0.0, 0.0, 0.0, 0.0, 0.0, 0.0, 0.0, 0.0, 0.0, 0.0, 0.0, 0.0, 0.0, 0.0, 0.0, 0.0, 0.0, 0.0, 0.0, 0.0, 0.0, 0.0, 0.0, 0.0, 0.0, 0.0, 0.0, 0.0, 0.0, 0.0, 0.0, 0.0, 0.0, 0.0, 0.0, 0.0, 0.0, 0.0, 0.0, 0.0, 0.0, 0.0, 0.0, 0.0, 0.0, 0.0, 0.0, 0.0, 0.0, 0.0, 0.0, 0.0, 0.0, 0.0, 0.0, 0.0, 0.0, 0.0, 0.0, 0.0, 0.0, 0.0, 0.0, 0.0, 0.0, 0.0, -0.0, -0.0, -0.0, -0.0, -0.0, -0.0, -0.0, -0.0, -0.0, -0.0, -0.0, -0.0, -0.0, -0.0, -0.0, -0.0, -0.0, -0.0, -0.0, -0.0, -0.0, -0.0, -0.0, -0.0, -0.0, -0.0, -0.0, -0.0, -0.0, -0.0, -0.0, -0.0, -0.0, -0.0, -0.0, -0.0, -0.0, -0.0, -0.0, -0.0, -0.0, -0.0, -0.0, -0.0, -0.0, -0.0, -0.0, -0.0, -0.0, -0.0, -0.0, -0.0, -0.0, -0.0, -0.0, -0.0, -0.0, -0.0, -0.0, -0.0, -0.0, -0.0, -0.0, -0.0, -0.0, -0.0, -0.0, -0.0, -0.0, -0.0, -1.7756006070928429E-5, -1.955926027849794E-5, -2.1265642444599059E-5, -2.2878087249309936E-5, -2.4399475238503513E-5, -2.5832632877734329E-5, -2.7180332648224444E-5, -2.8445293182983732E-5, -2.9630179441154765E-5, -3.0737602918726609E-5, -3.1770121893815045E-5, -3.2730241704758869E-5, -3.3620415059333691E-5, -3.4443042373434618E-5, -3.5200472137629193E-5, -3.5895001310030509E-5, -3.652887573398812E-5, -3.7104290579141277E-5, -3.7623390804425058E-5, -3.808827164166491E-5, -3.8500979098439383E-5, -3.886351047893401E-5, -3.9177814921551905E-5, -3.9445793952087749E-5, -3.966930205131298E-5, -3.98501472358593E-5, -3.9990091651326829E-5, -4.0090852176581095E-5, -4.0154101038240283E-5, -4.0181466434390562E-5, -4.017453316660271E-5, -4.013484327935801E-5, -4.0063896706025282E-5, -3.9963151920563813E-5, -3.9834026594159355E-5, -3.9677898256031791E-5, -3.9496104957683613E-5, -3.9289945939888413E-5, -3.9060682301747689E-5, -3.8809537671172525E-5, -3.8537698876174604E-5, -3.8246316616377579E-5, -3.793650613418646E-5, -3.7609347885077623E-5, -3.7265888206497395E-5, -3.6907139984880808E-5, -3.6534083320325723E-5, -3.6147666188480321E-5, -3.5748805099224027E-5, -3.5338385751743129E-5, 0.0, 0.0, 0.0, 0.0, 0.0, 0.0, 0.0, 0.0, 0.0, 0.0, 0.0, 0.0, 0.0, 0.0, 0.0, 0.0, 0.0, 0.0, 0.0, 0.0, 0.0, 0.0, 0.0, 0.0, 0.0, 0.0, 0.0, 0.0, 0.0, 0.0, 0.0, 0.0, 0.0, 0.0, 0.0, 0.0, 0.0, 0.0, 0.0, 0.0, 0.0, 0.0, 0.0, 0.0, 0.0, 0.0, 0.0, 0.0, 0.0, 0.0, 0.0, 0.0, 0.0, 0.0, 0.0, 0.0, 0.0, 0.0, 0.0, 0.0, 0.0, 0.0, 0.0, 0.0, 0.0, 0.0, 0.0, 0.0, 0.0, 0.0, 1.7756006070928429E-5, 1.955926027849794E-5, 2.1265642444599059E-5, 2.2878087249309936E-5, 2.4399475238503513E-5, 2.5832632877734329E-5, 2.7180332648224444E-5, 2.8445293182983732E-5, 2.9630179441154765E-5, 3.0737602918726609E-5, 3.1770121893815045E-5, 3.2730241704758869E-5, 3.3620415059333691E-5, 3.4443042373434618E-5, 3.5200472137629193E-5, 3.5895001310030509E-5, 3.652887573398812E-5, 3.7104290579141277E-5, 3.7623390804425058E-5, 3.808827164166491E-5, 3.8500979098439383E-5, 3.886351047893401E-5, 3.9177814921551905E-5, 3.9445793952087749E-5, 3.966930205131298E-5, 3.98501472358593E-5, 3.9990091651326829E-5, 4.0090852176581095E-5, 4.0154101038240283E-5, 4.0181466434390562E-5, 4.017453316660271E-5, 4.013484327935801E-5, 4.0063896706025282E-5, 3.9963151920563813E-5, 3.9834026594159355E-5, 3.9677898256031791E-5, 3.9496104957683613E-5, 3.9289945939888413E-5, 3.9060682301747689E-5, 3.8809537671172525E-5, 3.8537698876174604E-5, 3.8246316616377579E-5, 3.793650613418646E-5, 3.7609347885077623E-5, 3.7265888206497395E-5, 3.6907139984880808E-5, 3.6534083320325723E-5, 3.6147666188480321E-5, 3.5748805099224027E-5, 3.5338385751743129E-5, 0.0, 0.0, 0.0, 0.0, -0.0, -0.0, -0.0, -0.0, -0.0, -0.0, -0.0, -0.0, -0.0, -0.0, -0.0, -0.0, -0.0, -0.0, -0.0, -0.0, -0.0, -0.0, -0.0, -0.0, -0.0, -0.0, -0.0, -0.0, -0.0, -0.0, -0.0, -0.0, -0.0, -0.0, -0.0, -0.0, -0.0, -0.0, -0.0, -0.0, -0.0, -0.0, -0.0, -0.0, -0.0, -0.0, -0.0, -0.0, -0.0, -0.0, -0.0, -0.0, -0.0, -0.0, -0.0, -0.0, -0.0, -0.0, -0.0, -0.0, -0.0, -0.0, -0.0, -0.0, -0.0, -0.0, -0.0, -0.0, -0.0, -0.0, -0.0, -0.0, -0.0, -0.0, -0.0, -0.0, -0.0, -0.0, -0.0, -0.0, -0.0, -0.0, -0.0, -0.0, -0.0, -0.0, -0.0, -0.0, -0.0, -0.0, -0.0, -0.0, -0.0, -0.0, -0.0, -0.0, -0.0, -0.0, -0.0, -0.0, -0.0, -0.0, -0.0, -0.0, -0.0, -0.0, -0.0, -0.0, -0.0, -0.0, -0.0, -0.0, -0.0, -0.0, -0.0, -0.0, -0.0, -0.0, -0.0, -0.0, -0.0, -0.0, -0.0, -0.0, 0.0, 0.0, 0.0, 0.0, 0.0, 0.0, 0.0, 0.0, 0.0, 0.0, 0.0, 0.0, 0.0, 0.0, 0.0, 0.0, 0.0, 0.0, 0.0, 0.0, 0.0, 0.0, 0.0, 0.0, 0.0, 0.0, 0.0, 0.0, 0.0, 0.0, 0.0, 0.0, 0.0, 0.0, 0.0, 0.0, 0.0, 0.0, 0.0, 0.0, 0.0, 0.0, 0.0, 0.0, 0.0, 0.0, 0.0, 0.0, 0.0, 0.0, 0.0, 0.0, 0.0, 0.0, 0.0, 0.0, 0.0, 0.0, 0.0, 0.0, 0.0, 0.0, 0.0, 0.0, 0.0, 0.0, 0.0, 0.0, 0.0, 0.0, 0.0, 0.0, 0.0, 0.0, 0.0, 0.0, 0.0, 0.0, 0.0, 0.0, 0.0, 0.0, 0.0, 0.0, 0.0, 0.0, 0.0, 0.0, 0.0, 0.0, 0.0, 0.0, 0.0, 0.0, 0.0, 0.0, 0.0, 0.0, 0.0, 0.0, 0.0, 0.0, 0.0, 0.0, 0.0, 0.0, 0.0, 0.0, 0.0, 0.0, 0.0, 0.0, 0.0, 0.0, 0.0, 0.0, 0.0, 0.0, 0.0, 0.0, 0.0, 0.0, 0.0, 0.0, -0.0, -0.0, -0.0, -0.0, -0.0, -0.0, -0.0, -0.0, -0.0, -0.0, -0.0, -0.0, -0.0, -0.0, -0.0, -0.0, -0.0, -0.0, -0.0, -0.0, -0.0, -0.0, -0.0, -0.0, -0.0, -0.0, -0.0, -0.0, -0.0, -0.0, -0.0, -0.0, -0.0, -0.0, -0.0, -0.0, -0.0, -0.0, -0.0, -0.0, -0.0, -0.0, -0.0, -0.0, -0.0, -0.0, -0.0, -0.0, -0.0, -0.0, -0.0, -0.0, -0.0, -0.0, -0.0, -0.0, -0.0, -0.0, -0.0, -0.0, -0.0, -0.0, -0.0, -0.0, -0.0, -0.0, -0.0, -0.0, -0.0, -0.0, -0.0, -1.7756006070928429E-5, -1.955926027849794E-5, -2.1265642444599059E-5, -2.2878087249309936E-5, -2.4399475238503513E-5, -2.5832632877734329E-5, -2.7180332648224444E-5, -2.8445293182983732E-5, -2.9630179441154765E-5, -3.0737602918726609E-5, -3.1770121893815045E-5, -3.2730241704758869E-5, -3.3620415059333691E-5, -3.4443042373434618E-5, -3.5200472137629193E-5, -3.5895001310030509E-5, -3.652887573398812E-5, -3.7104290579141277E-5, -3.7623390804425058E-5, -3.808827164166491E-5, -3.8500979098439383E-5, -3.886351047893401E-5, -3.9177814921551905E-5, -3.9445793952087749E-5, -3.966930205131298E-5, -3.98501472358593E-5, -3.9990091651326829E-5, -4.0090852176581095E-5, -4.0154101038240283E-5, -4.0181466434390562E-5, -4.017453316660271E-5, -4.013484327935801E-5, -4.0063896706025282E-5, -3.9963151920563813E-5, -3.9834026594159355E-5, -3.9677898256031791E-5, -3.9496104957683613E-5, -3.9289945939888413E-5, -3.9060682301747689E-5, -3.8809537671172525E-5, -3.8537698876174604E-5, -3.8246316616377579E-5, -3.793650613418646E-5, -3.7609347885077623E-5, -3.7265888206497395E-5, -3.6907139984880808E-5, -3.6534083320325723E-5, -3.6147666188480321E-5, -3.5748805099224027E-5, 0.0, 0.0, 0.0, 0.0, 0.0, 0.0, 0.0, 0.0, 0.0, 0.0, 0.0, 0.0, 0.0, 0.0, 0.0, 0.0, 0.0, 0.0, 0.0, 0.0, 0.0, 0.0, 0.0, 0.0, 0.0, 0.0, 0.0, 0.0, 0.0, 0.0, 0.0, 0.0, 0.0, 0.0, 0.0, 0.0, 0.0, 0.0, 0.0, 0.0, 0.0, 0.0, 0.0, 0.0, 0.0, 0.0, 0.0, 0.0, 0.0, 0.0, 0.0, 0.0, 0.0, 0.0, 0.0, 0.0, 0.0, 0.0, 0.0, 0.0, 0.0, 0.0, 0.0, 0.0, 0.0, 0.0, 0.0, 0.0, 0.0, 0.0, 0.0, 1.7756006070928429E-5, 1.955926027849794E-5, 2.1265642444599059E-5, 2.2878087249309936E-5, 2.4399475238503513E-5, 2.5832632877734329E-5, 2.7180332648224444E-5, 2.8445293182983732E-5, 2.9630179441154765E-5, 3.0737602918726609E-5, 3.1770121893815045E-5, 3.2730241704758869E-5, 3.3620415059333691E-5, 3.4443042373434618E-5, 3.5200472137629193E-5, 3.5895001310030509E-5, 3.652887573398812E-5, 3.7104290579141277E-5, 3.7623390804425058E-5, 3.808827164166491E-5, 3.8500979098439383E-5, 3.886351047893401E-5, 3.9177814921551905E-5, 3.9445793952087749E-5, 3.966930205131298E-5, 3.98501472358593E-5, 3.9990091651326829E-5, 4.0090852176581095E-5, 4.0154101038240283E-5, 4.0181466434390562E-5, 4.017453316660271E-5, 4.013484327935801E-5, 4.0063896706025282E-5, 3.9963151920563813E-5, 3.9834026594159355E-5, 3.9677898256031791E-5, 3.9496104957683613E-5, 3.9289945939888413E-5, 3.9060682301747689E-5, 3.8809537671172525E-5, 3.8537698876174604E-5, 3.8246316616377579E-5, 3.793650613418646E-5, 3.7609347885077623E-5, 3.7265888206497395E-5, 3.6907139984880808E-5, 3.6534083320325723E-5, 3.6147666188480321E-5, 3.5748805099224027E-5, 0.0, 0.0, 0.0, 0.0, -0.0, -0.0, -0.0, -0.0, -0.0, -0.0, -0.0, -0.0, -0.0, -0.0, -0.0, -0.0, -0.0, -0.0, -0.0, -0.0, -0.0, -0.0, -0.0, -0.0, -0.0, -0.0, -0.0, -0.0, -0.0, -0.0, -0.0, -0.0, -0.0, -0.0, -0.0, -0.0, -0.0, -0.0, -0.0, -0.0, -0.0, -0.0, -0.0, -0.0, -0.0, -0.0, -0.0, -0.0, -0.0, -0.0, -0.0, -0.0, -0.0, -0.0, -0.0, -0.0, -0.0, -0.0, -0.0, -0.0, -0.0, -0.0, -0.0, -0.0, -0.0, -0.0, -0.0, -0.0, -0.0, -0.0, -0.0, -0.0, -0.0, -0.0, -0.0, -0.0, -0.0, -0.0, -0.0, -0.0, -0.0, -0.0, -0.0, -0.0, -0.0, -0.0, -0.0, -0.0, -0.0, -0.0, -0.0, -0.0, -0.0, -0.0, -0.0, -0.0, -0.0, -0.0, -0.0, -0.0, -0.0, -0.0, -0.0, -0.0, -0.0, -0.0, -0.0, -0.0, -0.0, -0.0, -0.0, -0.0, -0.0, -0.0, -0.0, -0.0, -0.0, -0.0, -0.0, -0.0, -0.0, -0.0, -0.0, -0.0, 0.0, 0.0, 0.0, 0.0, 0.0, 0.0, 0.0, 0.0, 0.0, 0.0, 0.0, 0.0, 0.0, 0.0, 0.0, 0.0, 0.0, 0.0, 0.0, 0.0, 0.0, 0.0, 0.0, 0.0, 0.0, 0.0, 0.0, 0.0, 0.0, 0.0, 0.0, 0.0, 0.0, 0.0, 0.0, 0.0, 0.0, 0.0, 0.0, 0.0, 0.0, 0.0, 0.0, 0.0, 0.0, 0.0, 0.0, 0.0, 0.0, 0.0, 0.0, 0.0, 0.0, 0.0, 0.0, 0.0, 0.0, 0.0, 0.0, 0.0, 0.0, 0.0, 0.0, 0.0, 0.0, 0.0, 0.0, 0.0, 0.0, 0.0, 0.0, 0.0, 0.0, 0.0, 0.0, 0.0, 0.0, 0.0, 0.0, 0.0, 0.0, 0.0, 0.0, 0.0, 0.0, 0.0, 0.0, 0.0, 0.0, 0.0, 0.0, 0.0, 0.0, 0.0, 0.0, 0.0, 0.0, 0.0, 0.0, 0.0, 0.0, 0.0, 0.0, 0.0, 0.0, 0.0, 0.0, 0.0, 0.0, 0.0, 0.0, 0.0, 0.0, 0.0, 0.0, 0.0, 0.0, 0.0, 0.0, 0.0, 0.0, 0.0, 0.0, 0.0, -0.0, -0.0, -0.0, -0.0, -0.0, -0.0, -0.0, -0.0, -0.0, -0.0, -0.0, -0.0, -0.0, -0.0, -0.0, -0.0, -0.0, -0.0, -0.0, -0.0, -0.0, -0.0, -0.0, -0.0, -0.0, -0.0, -0.0, -0.0, -0.0, -0.0, -0.0, -0.0, -0.0, -0.0, -0.0, -0.0, -0.0, -0.0, -0.0, -0.0, -0.0, -0.0, -0.0, -0.0, -0.0, -0.0, -0.0, -0.0, -0.0, -0.0, -0.0, -0.0, -0.0, -0.0, -0.0, -0.0, -0.0, -0.0, -0.0, -0.0, -0.0, -0.0, -0.0, -0.0, -0.0, -0.0, -0.0, -0.0, -0.0, -0.0, -0.0, -0.0, -1.7756006070928429E-5, -1.955926027849794E-5, -2.1265642444599059E-5, -2.2878087249309936E-5, -2.4399475238503513E-5, -2.5832632877734329E-5, -2.7180332648224444E-5, -2.8445293182983732E-5, -2.9630179441154765E-5, -3.0737602918726609E-5, -3.1770121893815045E-5, -3.2730241704758869E-5, -3.3620415059333691E-5, -3.4443042373434618E-5, -3.5200472137629193E-5, -3.5895001310030509E-5, -3.652887573398812E-5, -3.7104290579141277E-5, -3.7623390804425058E-5, -3.808827164166491E-5, -3.8500979098439383E-5, -3.886351047893401E-5, -3.9177814921551905E-5, -3.9445793952087749E-5, -3.966930205131298E-5, -3.98501472358593E-5, -3.9990091651326829E-5, -4.0090852176581095E-5, -4.0154101038240283E-5, -4.0181466434390562E-5, -4.017453316660271E-5, -4.013484327935801E-5, -4.0063896706025282E-5, -3.9963151920563813E-5, -3.9834026594159355E-5, -3.9677898256031791E-5, -3.9496104957683613E-5, -3.9289945939888413E-5, -3.9060682301747689E-5, -3.8809537671172525E-5, -3.8537698876174604E-5, -3.8246316616377579E-5, -3.793650613418646E-5, -3.7609347885077623E-5, -3.7265888206497395E-5, -3.6907139984880808E-5, -3.6534083320325723E-5, -3.6147666188480321E-5, 0.0, 0.0, 0.0, 0.0, 0.0, 0.0, 0.0, 0.0, 0.0, 0.0, 0.0, 0.0, 0.0, 0.0, 0.0, 0.0, 0.0, 0.0, 0.0, 0.0, 0.0, 0.0, 0.0, 0.0, 0.0, 0.0, 0.0, 0.0, 0.0, 0.0, 0.0, 0.0, 0.0, 0.0, 0.0, 0.0, 0.0, 0.0, 0.0, 0.0, 0.0, 0.0, 0.0, 0.0, 0.0, 0.0, 0.0, 0.0, 0.0, 0.0, 0.0, 0.0, 0.0, 0.0, 0.0, 0.0, 0.0, 0.0, 0.0, 0.0, 0.0, 0.0, 0.0, 0.0, 0.0, 0.0, 0.0, 0.0, 0.0, 0.0, 0.0, 0.0, 1.7756006070928429E-5, 1.955926027849794E-5, 2.1265642444599059E-5, 2.2878087249309936E-5, 2.4399475238503513E-5, 2.5832632877734329E-5, 2.7180332648224444E-5, 2.8445293182983732E-5, 2.9630179441154765E-5, 3.0737602918726609E-5, 3.1770121893815045E-5, 3.2730241704758869E-5, 3.3620415059333691E-5, 3.4443042373434618E-5, 3.5200472137629193E-5, 3.5895001310030509E-5, 3.652887573398812E-5, 3.7104290579141277E-5, 3.7623390804425058E-5, 3.808827164166491E-5, 3.8500979098439383E-5, 3.886351047893401E-5, 3.9177814921551905E-5, 3.9445793952087749E-5, 3.966930205131298E-5, 3.98501472358593E-5, 3.9990091651326829E-5, 4.0090852176581095E-5, 4.0154101038240283E-5, 4.0181466434390562E-5, 4.017453316660271E-5, 4.013484327935801E-5, 4.0063896706025282E-5, 3.9963151920563813E-5, 3.9834026594159355E-5, 3.9677898256031791E-5, 3.9496104957683613E-5, 3.9289945939888413E-5, 3.9060682301747689E-5, 3.8809537671172525E-5, 3.8537698876174604E-5, 3.8246316616377579E-5, 3.793650613418646E-5, 3.7609347885077623E-5, 3.7265888206497395E-5, 3.6907139984880808E-5, 3.6534083320325723E-5, 3.6147666188480321E-5, 0.0, 0.0, 0.0, 0.0, -0.0, -0.0, -0.0, -0.0, -0.0, -0.0, -0.0, -0.0, -0.0, -0.0, -0.0, -0.0, -0.0, -0.0, -0.0, -0.0, -0.0, -0.0, -0.0, -0.0, -0.0, -0.0, -0.0, -0.0, -0.0, -0.0, -0.0, -0.0, -0.0, -0.0, -0.0, -0.0, -0.0, -0.0, -0.0, -0.0, -0.0, -0.0, -0.0, -0.0, -0.0, -0.0, -0.0, -0.0, -0.0, -0.0, -0.0, -0.0, -0.0, -0.0, -0.0, -0.0, -0.0, -0.0, -0.0, -0.0, -0.0, -0.0, -0.0, -0.0, -0.0, -0.0, -0.0, -0.0, -0.0, -0.0, -0.0, -0.0, -0.0, -0.0, -0.0, -0.0, -0.0, -0.0, -0.0, -0.0, -0.0, -0.0, -0.0, -0.0, -0.0, -0.0, -0.0, -0.0, -0.0, -0.0, -0.0, -0.0, -0.0, -0.0, -0.0, -0.0, -0.0, -0.0, -0.0, -0.0, -0.0, -0.0, -0.0, -0.0, -0.0, -0.0, -0.0, -0.0, -0.0, -0.0, -0.0, -0.0, -0.0, -0.0, -0.0, -0.0, -0.0, -0.0, -0.0, -0.0, -0.0, -0.0, -0.0, -0.0, 0.0, 0.0, 0.0, 0.0, 0.0, 0.0, 0.0, 0.0, 0.0, 0.0, 0.0, 0.0, 0.0, 0.0, 0.0, 0.0, 0.0, 0.0, 0.0, 0.0, 0.0, 0.0, 0.0, 0.0, 0.0, 0.0, 0.0, 0.0, 0.0, 0.0, 0.0, 0.0, 0.0, 0.0, 0.0, 0.0, 0.0, 0.0, 0.0, 0.0, 0.0, 0.0, 0.0, 0.0, 0.0, 0.0, 0.0, 0.0, 0.0, 0.0, 0.0, 0.0, 0.0, 0.0, 0.0, 0.0, 0.0, 0.0, 0.0, 0.0, 0.0, 0.0, 0.0, 0.0, 0.0, 0.0, 0.0, 0.0, 0.0, 0.0, 0.0, 0.0, 0.0, 0.0, 0.0, 0.0, 0.0, 0.0, 0.0, 0.0, 0.0, 0.0, 0.0, 0.0, 0.0, 0.0, 0.0, 0.0, 0.0, 0.0, 0.0, 0.0, 0.0, 0.0, 0.0, 0.0, 0.0, 0.0, 0.0, 0.0, 0.0, 0.0, 0.0, 0.0, 0.0, 0.0, 0.0, 0.0, 0.0, 0.0, 0.0, 0.0, 0.0, 0.0, 0.0, 0.0, 0.0, 0.0, 0.0, 0.0, 0.0, 0.0, 0.0, 0.0, -0.0, -0.0, -0.0, -0.0, -0.0, -0.0, -0.0, -0.0, -0.0, -0.0, -0.0, -0.0, -0.0, -0.0, -0.0, -0.0, -0.0, -0.0, -0.0, -0.0, -0.0, -0.0, -0.0, -0.0, -0.0, -0.0, -0.0, -0.0, -0.0, -0.0, -0.0, -0.0, -0.0, -0.0, -0.0, -0.0, -0.0, -0.0, -0.0, -0.0, -0.0, -0.0, -0.0, -0.0, -0.0, -0.0, -0.0, -0.0, -0.0, -0.0, -0.0, -0.0, -0.0, -0.0, -0.0, -0.0, -0.0, -0.0, -0.0, -0.0, -0.0, -0.0, -0.0, -0.0, -0.0, -0.0, -0.0, -0.0, -0.0, -0.0, -0.0, -0.0, -0.0, -1.7756006070928429E-5, -1.955926027849794E-5, -2.1265642444599059E-5, -2.2878087249309936E-5, -2.4399475238503513E-5, -2.5832632877734329E-5, -2.7180332648224444E-5, -2.8445293182983732E-5, -2.9630179441154765E-5, -3.0737602918726609E-5, -3.1770121893815045E-5, -3.2730241704758869E-5, -3.3620415059333691E-5, -3.4443042373434618E-5, -3.5200472137629193E-5, -3.5895001310030509E-5, -3.652887573398812E-5, -3.7104290579141277E-5, -3.7623390804425058E-5, -3.808827164166491E-5, -3.8500979098439383E-5, -3.886351047893401E-5, -3.9177814921551905E-5, -3.9445793952087749E-5, -3.966930205131298E-5, -3.98501472358593E-5, -3.9990091651326829E-5, -4.0090852176581095E-5, -4.0154101038240283E-5, -4.0181466434390562E-5, -4.017453316660271E-5, -4.013484327935801E-5, -4.0063896706025282E-5, -3.9963151920563813E-5, -3.9834026594159355E-5, -3.9677898256031791E-5, -3.9496104957683613E-5, -3.9289945939888413E-5, -3.9060682301747689E-5, -3.8809537671172525E-5, -3.8537698876174604E-5, -3.8246316616377579E-5, -3.793650613418646E-5, -3.7609347885077623E-5, -3.7265888206497395E-5, -3.6907139984880808E-5, -3.6534083320325723E-5, 0.0, 0.0, 0.0, 0.0, 0.0, 0.0, 0.0, 0.0, 0.0, 0.0, 0.0, 0.0, 0.0, 0.0, 0.0, 0.0, 0.0, 0.0, 0.0, 0.0, 0.0, 0.0, 0.0, 0.0, 0.0, 0.0, 0.0, 0.0, 0.0, 0.0, 0.0, 0.0, 0.0, 0.0, 0.0, 0.0, 0.0, 0.0, 0.0, 0.0, 0.0, 0.0, 0.0, 0.0, 0.0, 0.0, 0.0, 0.0, 0.0, 0.0, 0.0, 0.0, 0.0, 0.0, 0.0, 0.0, 0.0, 0.0, 0.0, 0.0, 0.0, 0.0, 0.0, 0.0, 0.0, 0.0, 0.0, 0.0, 0.0, 0.0, 0.0, 0.0, 0.0, 1.7756006070928429E-5, 1.955926027849794E-5, 2.1265642444599059E-5, 2.2878087249309936E-5, 2.4399475238503513E-5, 2.5832632877734329E-5, 2.7180332648224444E-5, 2.8445293182983732E-5, 2.9630179441154765E-5, 3.0737602918726609E-5, 3.1770121893815045E-5, 3.2730241704758869E-5, 3.3620415059333691E-5, 3.4443042373434618E-5, 3.5200472137629193E-5, 3.5895001310030509E-5, 3.652887573398812E-5, 3.7104290579141277E-5, 3.7623390804425058E-5, 3.808827164166491E-5, 3.8500979098439383E-5, 3.886351047893401E-5, 3.9177814921551905E-5, 3.9445793952087749E-5, 3.966930205131298E-5, 3.98501472358593E-5, 3.9990091651326829E-5, 4.0090852176581095E-5, 4.0154101038240283E-5, 4.0181466434390562E-5, 4.017453316660271E-5, 4.013484327935801E-5, 4.0063896706025282E-5, 3.9963151920563813E-5, 3.9834026594159355E-5, 3.9677898256031791E-5, 3.9496104957683613E-5, 3.9289945939888413E-5, 3.9060682301747689E-5, 3.8809537671172525E-5, 3.8537698876174604E-5, 3.8246316616377579E-5, 3.793650613418646E-5, 3.7609347885077623E-5, 3.7265888206497395E-5, 3.6907139984880808E-5, 3.6534083320325723E-5, 0.0, 0.0, 0.0, 0.0, -0.0, -0.0, -0.0, -0.0, -0.0, -0.0, -0.0, -0.0, -0.0, -0.0, -0.0, -0.0, -0.0, -0.0, -0.0, -0.0, -0.0, -0.0, -0.0, -0.0, -0.0, -0.0, -0.0, -0.0, -0.0, -0.0, -0.0, -0.0, -0.0, -0.0, -0.0, -0.0, -0.0, -0.0, -0.0, -0.0, -0.0, -0.0, -0.0, -0.0, -0.0, -0.0, -0.0, -0.0, -0.0, -0.0, -0.0, -0.0, -0.0, -0.0, -0.0, -0.0, -0.0, -0.0, -0.0, -0.0, -0.0, -0.0, -0.0, -0.0, -0.0, -0.0, -0.0, -0.0, -0.0, -0.0, -0.0, -0.0, -0.0, -0.0, -0.0, -0.0, -0.0, -0.0, -0.0, -0.0, -0.0, -0.0, -0.0, -0.0, -0.0, -0.0, -0.0, -0.0, -0.0, -0.0, -0.0, -0.0, -0.0, -0.0, -0.0, -0.0, -0.0, -0.0, -0.0, -0.0, -0.0, -0.0, -0.0, -0.0, -0.0, -0.0, -0.0, -0.0, -0.0, -0.0, -0.0, -0.0, -0.0, -0.0, -0.0, -0.0, -0.0, -0.0, -0.0, -0.0, -0.0, -0.0, -0.0, -0.0, 0.0, 0.0, 0.0, 0.0, 0.0, 0.0, 0.0, 0.0, 0.0, 0.0, 0.0, 0.0, 0.0, 0.0, 0.0, 0.0, 0.0, 0.0, 0.0, 0.0, 0.0, 0.0, 0.0, 0.0, 0.0, 0.0, 0.0, 0.0, 0.0, 0.0, 0.0, 0.0, 0.0, 0.0, 0.0, 0.0, 0.0, 0.0, 0.0, 0.0, 0.0, 0.0, 0.0, 0.0, 0.0, 0.0, 0.0, 0.0, 0.0, 0.0, 0.0, 0.0, 0.0, 0.0, 0.0, 0.0, 0.0, 0.0, 0.0, 0.0, 0.0, 0.0, 0.0, 0.0, 0.0, 0.0, 0.0, 0.0, 0.0, 0.0, 0.0, 0.0, 0.0, 0.0, 0.0, 0.0, 0.0, 0.0, 0.0, 0.0, 0.0, 0.0, 0.0, 0.0, 0.0, 0.0, 0.0, 0.0, 0.0, 0.0, 0.0, 0.0, 0.0, 0.0, 0.0, 0.0, 0.0, 0.0, 0.0, 0.0, 0.0, 0.0, 0.0, 0.0, 0.0, 0.0, 0.0, 0.0, 0.0, 0.0, 0.0, 0.0, 0.0, 0.0, 0.0, 0.0, 0.0, 0.0, 0.0, 0.0, 0.0, 0.0, 0.0, 0.0, -0.0, -0.0, -0.0, -0.0, -0.0, -0.0, -0.0, -0.0, -0.0, -0.0, -0.0, -0.0, -0.0, -0.0, -0.0, -0.0, -0.0, -0.0, -0.0, -0.0, -0.0, -0.0, -0.0, -0.0, -0.0, -0.0, -0.0, -0.0, -0.0, -0.0, -0.0, -0.0, -0.0, -0.0, -0.0, -0.0, -0.0, -0.0, -0.0, -0.0, -0.0, -0.0, -0.0, -0.0, -0.0, -0.0, -0.0, -0.0, -0.0, -0.0, -0.0, -0.0, -0.0, -0.0, -0.0, -0.0, -0.0, -0.0, -0.0, -0.0, -0.0, -0.0, -0.0, -0.0, -0.0, -0.0, -0.0, -0.0, -0.0, -0.0, -0.0, -0.0, -0.0, -0.0, -1.7756006070928429E-5, -1.955926027849794E-5, -2.1265642444599059E-5, -2.2878087249309936E-5, -2.4399475238503513E-5, -2.5832632877734329E-5, -2.7180332648224444E-5, -2.8445293182983732E-5, -2.9630179441154765E-5, -3.0737602918726609E-5, -3.1770121893815045E-5, -3.2730241704758869E-5, -3.3620415059333691E-5, -3.4443042373434618E-5, -3.5200472137629193E-5, -3.5895001310030509E-5, -3.652887573398812E-5, -3.7104290579141277E-5, -3.7623390804425058E-5, -3.808827164166491E-5, -3.8500979098439383E-5, -3.886351047893401E-5, -3.9177814921551905E-5, -3.9445793952087749E-5, -3.966930205131298E-5, -3.98501472358593E-5, -3.9990091651326829E-5, -4.0090852176581095E-5, -4.0154101038240283E-5, -4.0181466434390562E-5, -4.017453316660271E-5, -4.013484327935801E-5, -4.0063896706025282E-5, -3.9963151920563813E-5, -3.9834026594159355E-5, -3.9677898256031791E-5, -3.9496104957683613E-5, -3.9289945939888413E-5, -3.9060682301747689E-5, -3.8809537671172525E-5, -3.8537698876174604E-5, -3.8246316616377579E-5, -3.793650613418646E-5, -3.7609347885077623E-5, -3.7265888206497395E-5, -3.6907139984880808E-5, 0.0, 0.0, 0.0, 0.0, 0.0, 0.0, 0.0, 0.0, 0.0, 0.0, 0.0, 0.0, 0.0, 0.0, 0.0, 0.0, 0.0, 0.0, 0.0, 0.0, 0.0, 0.0, 0.0, 0.0, 0.0, 0.0, 0.0, 0.0, 0.0, 0.0, 0.0, 0.0, 0.0, 0.0, 0.0, 0.0, 0.0, 0.0, 0.0, 0.0, 0.0, 0.0, 0.0, 0.0, 0.0, 0.0, 0.0, 0.0, 0.0, 0.0, 0.0, 0.0, 0.0, 0.0, 0.0, 0.0, 0.0, 0.0, 0.0, 0.0, 0.0, 0.0, 0.0, 0.0, 0.0, 0.0, 0.0, 0.0, 0.0, 0.0, 0.0, 0.0, 0.0, 0.0, 1.7756006070928429E-5, 1.955926027849794E-5, 2.1265642444599059E-5, 2.2878087249309936E-5, 2.4399475238503513E-5, 2.5832632877734329E-5, 2.7180332648224444E-5, 2.8445293182983732E-5, 2.9630179441154765E-5, 3.0737602918726609E-5, 3.1770121893815045E-5, 3.2730241704758869E-5, 3.3620415059333691E-5, 3.4443042373434618E-5, 3.5200472137629193E-5, 3.5895001310030509E-5, 3.652887573398812E-5, 3.7104290579141277E-5, 3.7623390804425058E-5, 3.808827164166491E-5, 3.8500979098439383E-5, 3.886351047893401E-5, 3.9177814921551905E-5, 3.9445793952087749E-5, 3.966930205131298E-5, 3.98501472358593E-5, 3.9990091651326829E-5, 4.0090852176581095E-5, 4.0154101038240283E-5, 4.0181466434390562E-5, 4.017453316660271E-5, 4.013484327935801E-5, 4.0063896706025282E-5, 3.9963151920563813E-5, 3.9834026594159355E-5, 3.9677898256031791E-5, 3.9496104957683613E-5, 3.9289945939888413E-5, 3.9060682301747689E-5, 3.8809537671172525E-5, 3.8537698876174604E-5, 3.8246316616377579E-5, 3.793650613418646E-5, 3.7609347885077623E-5, 3.7265888206497395E-5, 3.6907139984880808E-5, 0.0, 0.0, 0.0, 0.0, -0.0, -0.0, -0.0, -0.0, -0.0, -0.0, -0.0, -0.0, -0.0, -0.0, -0.0, -0.0, -0.0, -0.0, -0.0, -0.0, -0.0, -0.0, -0.0, -0.0, -0.0, -0.0, -0.0, -0.0, -0.0, -0.0, -0.0, -0.0, -0.0, -0.0, -0.0, -0.0, -0.0, -0.0, -0.0, -0.0, -0.0, -0.0, -0.0, -0.0, -0.0, -0.0, -0.0, -0.0, -0.0, -0.0, -0.0, -0.0, -0.0, -0.0, -0.0, -0.0, -0.0, -0.0, -0.0, -0.0, -0.0, -0.0, -0.0, -0.0, -0.0, -0.0, -0.0, -0.0, -0.0, -0.0, -0.0, -0.0, -0.0, -0.0, -0.0, -0.0, -0.0, -0.0, -0.0, -0.0, -0.0, -0.0, -0.0, -0.0, -0.0, -0.0, -0.0, -0.0, -0.0, -0.0, -0.0, -0.0, -0.0, -0.0, -0.0, -0.0, -0.0, -0.0, -0.0, -0.0, -0.0, -0.0, -0.0, -0.0, -0.0, -0.0, -0.0, -0.0, -0.0, -0.0, -0.0, -0.0, -0.0, -0.0, -0.0, -0.0, -0.0, -0.0, -0.0, -0.0, -0.0, -0.0, -0.0, -0.0, 0.0, 0.0, 0.0, 0.0, 0.0, 0.0, 0.0, 0.0, 0.0, 0.0, 0.0, 0.0, 0.0, 0.0, 0.0, 0.0, 0.0, 0.0, 0.0, 0.0, 0.0, 0.0, 0.0, 0.0, 0.0, 0.0, 0.0, 0.0, 0.0, 0.0, 0.0, 0.0, 0.0, 0.0, 0.0, 0.0, 0.0, 0.0, 0.0, 0.0, 0.0, 0.0, 0.0, 0.0, 0.0, 0.0, 0.0, 0.0, 0.0, 0.0, 0.0, 0.0, 0.0, 0.0, 0.0, 0.0, 0.0, 0.0, 0.0, 0.0, 0.0, 0.0, 0.0, 0.0, 0.0, 0.0, 0.0, 0.0, 0.0, 0.0, 0.0, 0.0, 0.0, 0.0, 0.0, 0.0, 0.0, 0.0, 0.0, 0.0, 0.0, 0.0, 0.0, 0.0, 0.0, 0.0, 0.0, 0.0, 0.0, 0.0, 0.0, 0.0, 0.0, 0.0, 0.0, 0.0, 0.0, 0.0, 0.0, 0.0, 0.0, 0.0, 0.0, 0.0, 0.0, 0.0, 0.0, 0.0, 0.0, 0.0, 0.0, 0.0, 0.0, 0.0, 0.0, 0.0, 0.0, 0.0, 0.0, 0.0, 0.0, 0.0, 0.0, 0.0, -0.0, -0.0, -0.0, -0.0, -0.0, -0.0, -0.0, -0.0, -0.0, -0.0, -0.0, -0.0, -0.0, -0.0, -0.0, -0.0, -0.0, -0.0, -0.0, -0.0, -0.0, -0.0, -0.0, -0.0, -0.0, -0.0, -0.0, -0.0, -0.0, -0.0, -0.0, -0.0, -0.0, -0.0, -0.0, -0.0, -0.0, -0.0, -0.0, -0.0, -0.0, -0.0, -0.0, -0.0, -0.0, -0.0, -0.0, -0.0, -0.0, -0.0, -0.0, -0.0, -0.0, -0.0, -0.0, -0.0, -0.0, -0.0, -0.0, -0.0, -0.0, -0.0, -0.0, -0.0, -0.0, -0.0, -0.0, -0.0, -0.0, -0.0, -0.0, -0.0, -0.0, -0.0, -0.0, -1.7756006070928429E-5, -1.955926027849794E-5, -2.1265642444599059E-5, -2.2878087249309936E-5, -2.4399475238503513E-5, -2.5832632877734329E-5, -2.7180332648224444E-5, -2.8445293182983732E-5, -2.9630179441154765E-5, -3.0737602918726609E-5, -3.1770121893815045E-5, -3.2730241704758869E-5, -3.3620415059333691E-5, -3.4443042373434618E-5, -3.5200472137629193E-5, -3.5895001310030509E-5, -3.652887573398812E-5, -3.7104290579141277E-5, -3.7623390804425058E-5, -3.808827164166491E-5, -3.8500979098439383E-5, -3.886351047893401E-5, -3.9177814921551905E-5, -3.9445793952087749E-5, -3.966930205131298E-5, -3.98501472358593E-5, -3.9990091651326829E-5, -4.0090852176581095E-5, -4.0154101038240283E-5, -4.0181466434390562E-5, -4.017453316660271E-5, -4.013484327935801E-5, -4.0063896706025282E-5, -3.9963151920563813E-5, -3.9834026594159355E-5, -3.9677898256031791E-5, -3.9496104957683613E-5, -3.9289945939888413E-5, -3.9060682301747689E-5, -3.8809537671172525E-5, -3.8537698876174604E-5, -3.8246316616377579E-5, -3.793650613418646E-5, -3.7609347885077623E-5, -3.7265888206497395E-5, 0.0, 0.0, 0.0, 0.0, 0.0, 0.0, 0.0, 0.0, 0.0, 0.0, 0.0, 0.0, 0.0, 0.0, 0.0, 0.0, 0.0, 0.0, 0.0, 0.0, 0.0, 0.0, 0.0, 0.0, 0.0, 0.0, 0.0, 0.0, 0.0, 0.0, 0.0, 0.0, 0.0, 0.0, 0.0, 0.0, 0.0, 0.0, 0.0, 0.0, 0.0, 0.0, 0.0, 0.0, 0.0, 0.0, 0.0, 0.0, 0.0, 0.0, 0.0, 0.0, 0.0, 0.0, 0.0, 0.0, 0.0, 0.0, 0.0, 0.0, 0.0, 0.0, 0.0, 0.0, 0.0, 0.0, 0.0, 0.0, 0.0, 0.0, 0.0, 0.0, 0.0, 0.0, 0.0, 1.7756006070928429E-5, 1.955926027849794E-5, 2.1265642444599059E-5, 2.2878087249309936E-5, 2.4399475238503513E-5, 2.5832632877734329E-5, 2.7180332648224444E-5, 2.8445293182983732E-5, 2.9630179441154765E-5, 3.0737602918726609E-5, 3.1770121893815045E-5, 3.2730241704758869E-5, 3.3620415059333691E-5, 3.4443042373434618E-5, 3.5200472137629193E-5, 3.5895001310030509E-5, 3.652887573398812E-5, 3.7104290579141277E-5, 3.7623390804425058E-5, 3.808827164166491E-5, 3.8500979098439383E-5, 3.886351047893401E-5, 3.9177814921551905E-5, 3.9445793952087749E-5, 3.966930205131298E-5, 3.98501472358593E-5, 3.9990091651326829E-5, 4.0090852176581095E-5, 4.0154101038240283E-5, 4.0181466434390562E-5, 4.017453316660271E-5, 4.013484327935801E-5, 4.0063896706025282E-5, 3.9963151920563813E-5, 3.9834026594159355E-5, 3.9677898256031791E-5, 3.9496104957683613E-5, 3.9289945939888413E-5, 3.9060682301747689E-5, 3.8809537671172525E-5, 3.8537698876174604E-5, 3.8246316616377579E-5, 3.793650613418646E-5, 3.7609347885077623E-5, 3.7265888206497395E-5, 0.0, 0.0, 0.0, 0.0, -0.0, -0.0, -0.0, -0.0, -0.0, -0.0, -0.0, -0.0, -0.0, -0.0, -0.0, -0.0, -0.0, -0.0, -0.0, -0.0, -0.0, -0.0, -0.0, -0.0, -0.0, -0.0, -0.0, -0.0, -0.0, -0.0, -0.0, -0.0, -0.0, -0.0, -0.0, -0.0, -0.0, -0.0, -0.0, -0.0, -0.0, -0.0, -0.0, -0.0, -0.0, -0.0, -0.0, -0.0, -0.0, -0.0, -0.0, -0.0, -0.0, -0.0, -0.0, -0.0, -0.0, -0.0, -0.0, -0.0, -0.0, -0.0, -0.0, -0.0, -0.0, -0.0, -0.0, -0.0, -0.0, -0.0, -0.0, -0.0, -0.0, -0.0, -0.0, -0.0, -0.0, -0.0, -0.0, -0.0, -0.0, -0.0, -0.0, -0.0, -0.0, -0.0, -0.0, -0.0, -0.0, -0.0, -0.0, -0.0, -0.0, -0.0, -0.0, -0.0, -0.0, -0.0, -0.0, -0.0, -0.0, -0.0, -0.0, -0.0, -0.0, -0.0, -0.0, -0.0, -0.0, -0.0, -0.0, -0.0, -0.0, -0.0, -0.0, -0.0, -0.0, -0.0, -0.0, -0.0, -0.0, -0.0, -0.0, -0.0, 0.0, 0.0, 0.0, 0.0, 0.0, 0.0, 0.0, 0.0, 0.0, 0.0, 0.0, 0.0, 0.0, 0.0, 0.0, 0.0, 0.0, 0.0, 0.0, 0.0, 0.0, 0.0, 0.0, 0.0, 0.0, 0.0, 0.0, 0.0, 0.0, 0.0, 0.0, 0.0, 0.0, 0.0, 0.0, 0.0, 0.0, 0.0, 0.0, 0.0, 0.0, 0.0, 0.0, 0.0, 0.0, 0.0, 0.0, 0.0, 0.0, 0.0, 0.0, 0.0, 0.0, 0.0, 0.0, 0.0, 0.0, 0.0, 0.0, 0.0, 0.0, 0.0, 0.0, 0.0, 0.0, 0.0, 0.0, 0.0, 0.0, 0.0, 0.0, 0.0, 0.0, 0.0, 0.0, 0.0, 0.0, 0.0, 0.0, 0.0, 0.0, 0.0, 0.0, 0.0, 0.0, 0.0, 0.0, 0.0, 0.0, 0.0, 0.0, 0.0, 0.0, 0.0, 0.0, 0.0, 0.0, 0.0, 0.0, 0.0, 0.0, 0.0, 0.0, 0.0, 0.0, 0.0, 0.0, 0.0, 0.0, 0.0, 0.0, 0.0, 0.0, 0.0, 0.0, 0.0, 0.0, 0.0, 0.0, 0.0, 0.0, 0.0, 0.0, 0.0, -0.0, -0.0, -0.0, -0.0, -0.0, -0.0, -0.0, -0.0, -0.0, -0.0, -0.0, -0.0, -0.0, -0.0, -0.0, -0.0, -0.0, -0.0, -0.0, -0.0, -0.0, -0.0, -0.0, -0.0, -0.0, -0.0, -0.0, -0.0, -0.0, -0.0, -0.0, -0.0, -0.0, -0.0, -0.0, -0.0, -0.0, -0.0, -0.0, -0.0, -0.0, -0.0, -0.0, -0.0, -0.0, -0.0, -0.0, -0.0, -0.0, -0.0, -0.0, -0.0, -0.0, -0.0, -0.0, -0.0, -0.0, -0.0, -0.0, -0.0, -0.0, -0.0, -0.0, -0.0, -0.0, -0.0, -0.0, -0.0, -0.0, -0.0, -0.0, -0.0, -0.0, -0.0, -0.0, -0.0, -1.7756006070928429E-5, -1.955926027849794E-5, -2.1265642444599059E-5, -2.2878087249309936E-5, -2.4399475238503513E-5, -2.5832632877734329E-5, -2.7180332648224444E-5, -2.8445293182983732E-5, -2.9630179441154765E-5, -3.0737602918726609E-5, -3.1770121893815045E-5, -3.2730241704758869E-5, -3.3620415059333691E-5, -3.4443042373434618E-5, -3.5200472137629193E-5, -3.5895001310030509E-5, -3.652887573398812E-5, -3.7104290579141277E-5, -3.7623390804425058E-5, -3.808827164166491E-5, -3.8500979098439383E-5, -3.886351047893401E-5, -3.9177814921551905E-5, -3.9445793952087749E-5, -3.966930205131298E-5, -3.98501472358593E-5, -3.9990091651326829E-5, -4.0090852176581095E-5, -4.0154101038240283E-5, -4.0181466434390562E-5, -4.017453316660271E-5, -4.013484327935801E-5, -4.0063896706025282E-5, -3.9963151920563813E-5, -3.9834026594159355E-5, -3.9677898256031791E-5, -3.9496104957683613E-5, -3.9289945939888413E-5, -3.9060682301747689E-5, -3.8809537671172525E-5, -3.8537698876174604E-5, -3.8246316616377579E-5, -3.793650613418646E-5, -3.7609347885077623E-5, 0.0, 0.0, 0.0, 0.0, 0.0, 0.0, 0.0, 0.0, 0.0, 0.0, 0.0, 0.0, 0.0, 0.0, 0.0, 0.0, 0.0, 0.0, 0.0, 0.0, 0.0, 0.0, 0.0, 0.0, 0.0, 0.0, 0.0, 0.0, 0.0, 0.0, 0.0, 0.0, 0.0, 0.0, 0.0, 0.0, 0.0, 0.0, 0.0, 0.0, 0.0, 0.0, 0.0, 0.0, 0.0, 0.0, 0.0, 0.0, 0.0, 0.0, 0.0, 0.0, 0.0, 0.0, 0.0, 0.0, 0.0, 0.0, 0.0, 0.0, 0.0, 0.0, 0.0, 0.0, 0.0, 0.0, 0.0, 0.0, 0.0, 0.0, 0.0, 0.0, 0.0, 0.0, 0.0, 0.0, 1.7756006070928429E-5, 1.955926027849794E-5, 2.1265642444599059E-5, 2.2878087249309936E-5, 2.4399475238503513E-5, 2.5832632877734329E-5, 2.7180332648224444E-5, 2.8445293182983732E-5, 2.9630179441154765E-5, 3.0737602918726609E-5, 3.1770121893815045E-5, 3.2730241704758869E-5, 3.3620415059333691E-5, 3.4443042373434618E-5, 3.5200472137629193E-5, 3.5895001310030509E-5, 3.652887573398812E-5, 3.7104290579141277E-5, 3.7623390804425058E-5, 3.808827164166491E-5, 3.8500979098439383E-5, 3.886351047893401E-5, 3.9177814921551905E-5, 3.9445793952087749E-5, 3.966930205131298E-5, 3.98501472358593E-5, 3.9990091651326829E-5, 4.0090852176581095E-5, 4.0154101038240283E-5, 4.0181466434390562E-5, 4.017453316660271E-5, 4.013484327935801E-5, 4.0063896706025282E-5, 3.9963151920563813E-5, 3.9834026594159355E-5, 3.9677898256031791E-5, 3.9496104957683613E-5, 3.9289945939888413E-5, 3.9060682301747689E-5, 3.8809537671172525E-5, 3.8537698876174604E-5, 3.8246316616377579E-5, 3.793650613418646E-5, 3.7609347885077623E-5, 0.0, 0.0, 0.0, 0.0, -0.0, -0.0, -0.0, -0.0, -0.0, -0.0, -0.0, -0.0, -0.0, -0.0, -0.0, -0.0, -0.0, -0.0, -0.0, -0.0, -0.0, -0.0, -0.0, -0.0, -0.0, -0.0, -0.0, -0.0, -0.0, -0.0, -0.0, -0.0, -0.0, -0.0, -0.0, -0.0, -0.0, -0.0, -0.0, -0.0, -0.0, -0.0, -0.0, -0.0, -0.0, -0.0, -0.0, -0.0, -0.0, -0.0, -0.0, -0.0, -0.0, -0.0, -0.0, -0.0, -0.0, -0.0, -0.0, -0.0, -0.0, -0.0, -0.0, -0.0, -0.0, -0.0, -0.0, -0.0, -0.0, -0.0, -0.0, -0.0, -0.0, -0.0, -0.0, -0.0, -0.0, -0.0, -0.0, -0.0, -0.0, -0.0, -0.0, -0.0, -0.0, -0.0, -0.0, -0.0, -0.0, -0.0, -0.0, -0.0, -0.0, -0.0, -0.0, -0.0, -0.0, -0.0, -0.0, -0.0, -0.0, -0.0, -0.0, -0.0, -0.0, -0.0, -0.0, -0.0, -0.0, -0.0, -0.0, -0.0, -0.0, -0.0, -0.0, -0.0, -0.0, -0.0, -0.0, -0.0, -0.0, -0.0, -0.0, -0.0, 0.0, 0.0, 0.0, 0.0, 0.0, 0.0, 0.0, 0.0, 0.0, 0.0, 0.0, 0.0, 0.0, 0.0, 0.0, 0.0, 0.0, 0.0, 0.0, 0.0, 0.0, 0.0, 0.0, 0.0, 0.0, 0.0, 0.0, 0.0, 0.0, 0.0, 0.0, 0.0, 0.0, 0.0, 0.0, 0.0, 0.0, 0.0, 0.0, 0.0, 0.0, 0.0, 0.0, 0.0, 0.0, 0.0, 0.0, 0.0, 0.0, 0.0, 0.0, 0.0, 0.0, 0.0, 0.0, 0.0, 0.0, 0.0, 0.0, 0.0, 0.0, 0.0, 0.0, 0.0, 0.0, 0.0, 0.0, 0.0, 0.0, 0.0, 0.0, 0.0, 0.0, 0.0, 0.0, 0.0, 0.0, 0.0, 0.0, 0.0, 0.0, 0.0, 0.0, 0.0, 0.0, 0.0, 0.0, 0.0, 0.0, 0.0, 0.0, 0.0, 0.0, 0.0, 0.0, 0.0, 0.0, 0.0, 0.0, 0.0, 0.0, 0.0, 0.0, 0.0, 0.0, 0.0, 0.0, 0.0, 0.0, 0.0, 0.0, 0.0, 0.0, 0.0, 0.0, 0.0, 0.0, 0.0, 0.0, 0.0, 0.0, 0.0, 0.0, 0.0, -0.0, -0.0, -0.0, -0.0, -0.0, -0.0, -0.0, -0.0, -0.0, -0.0, -0.0, -0.0, -0.0, -0.0, -0.0, -0.0, -0.0, -0.0, -0.0, -0.0, -0.0, -0.0, -0.0, -0.0, -0.0, -0.0, -0.0, -0.0, -0.0, -0.0, -0.0, -0.0, -0.0, -0.0, -0.0, -0.0, -0.0, -0.0, -0.0, -0.0, -0.0, -0.0, -0.0, -0.0, -0.0, -0.0, -0.0, -0.0, -0.0, -0.0, -0.0, -0.0, -0.0, -0.0, -0.0, -0.0, -0.0, -0.0, -0.0, -0.0, -0.0, -0.0, -0.0, -0.0, -0.0, -0.0, -0.0, -0.0, -0.0, -0.0, -0.0, -0.0, -0.0, -0.0, -0.0, -0.0, -0.0, -1.7756006070928429E-5, -1.955926027849794E-5, -2.1265642444599059E-5, -2.2878087249309936E-5, -2.4399475238503513E-5, -2.5832632877734329E-5, -2.7180332648224444E-5, -2.8445293182983732E-5, -2.9630179441154765E-5, -3.0737602918726609E-5, -3.1770121893815045E-5, -3.2730241704758869E-5, -3.3620415059333691E-5, -3.4443042373434618E-5, -3.5200472137629193E-5, -3.5895001310030509E-5, -3.652887573398812E-5, -3.7104290579141277E-5, -3.7623390804425058E-5, -3.808827164166491E-5, -3.8500979098439383E-5, -3.886351047893401E-5, -3.9177814921551905E-5, -3.9445793952087749E-5, -3.966930205131298E-5, -3.98501472358593E-5, -3.9990091651326829E-5, -4.0090852176581095E-5, -4.0154101038240283E-5, -4.0181466434390562E-5, -4.017453316660271E-5, -4.013484327935801E-5, -4.0063896706025282E-5, -3.9963151920563813E-5, -3.9834026594159355E-5, -3.9677898256031791E-5, -3.9496104957683613E-5, -3.9289945939888413E-5, -3.9060682301747689E-5, -3.8809537671172525E-5, -3.8537698876174604E-5, -3.8246316616377579E-5, -3.793650613418646E-5, 0.0, 0.0, 0.0, 0.0, 0.0, 0.0, 0.0, 0.0, 0.0, 0.0, 0.0, 0.0, 0.0, 0.0, 0.0, 0.0, 0.0, 0.0, 0.0, 0.0, 0.0, 0.0, 0.0, 0.0, 0.0, 0.0, 0.0, 0.0, 0.0, 0.0, 0.0, 0.0, 0.0, 0.0, 0.0, 0.0, 0.0, 0.0, 0.0, 0.0, 0.0, 0.0, 0.0, 0.0, 0.0, 0.0, 0.0, 0.0, 0.0, 0.0, 0.0, 0.0, 0.0, 0.0, 0.0, 0.0, 0.0, 0.0, 0.0, 0.0, 0.0, 0.0, 0.0, 0.0, 0.0, 0.0, 0.0, 0.0, 0.0, 0.0, 0.0, 0.0, 0.0, 0.0, 0.0, 0.0, 0.0, 1.7756006070928429E-5, 1.955926027849794E-5, 2.1265642444599059E-5, 2.2878087249309936E-5, 2.4399475238503513E-5, 2.5832632877734329E-5, 2.7180332648224444E-5, 2.8445293182983732E-5, 2.9630179441154765E-5, 3.0737602918726609E-5, 3.1770121893815045E-5, 3.2730241704758869E-5, 3.3620415059333691E-5, 3.4443042373434618E-5, 3.5200472137629193E-5, 3.5895001310030509E-5, 3.652887573398812E-5, 3.7104290579141277E-5, 3.7623390804425058E-5, 3.808827164166491E-5, 3.8500979098439383E-5, 3.886351047893401E-5, 3.9177814921551905E-5, 3.9445793952087749E-5, 3.966930205131298E-5, 3.98501472358593E-5, 3.9990091651326829E-5, 4.0090852176581095E-5, 4.0154101038240283E-5, 4.0181466434390562E-5, 4.017453316660271E-5, 4.013484327935801E-5, 4.0063896706025282E-5, 3.9963151920563813E-5, 3.9834026594159355E-5, 3.9677898256031791E-5, 3.9496104957683613E-5, 3.9289945939888413E-5, 3.9060682301747689E-5, 3.8809537671172525E-5, 3.8537698876174604E-5, 3.8246316616377579E-5, 3.793650613418646E-5, 0.0, 0.0, 0.0, 0.0, -0.0, -0.0, -0.0, -0.0, -0.0, -0.0, -0.0, -0.0, -0.0, -0.0, -0.0, -0.0, -0.0, -0.0, -0.0, -0.0, -0.0, -0.0, -0.0, -0.0, -0.0, -0.0, -0.0, -0.0, -0.0, -0.0, -0.0, -0.0, -0.0, -0.0, -0.0, -0.0, -0.0, -0.0, -0.0, -0.0, -0.0, -0.0, -0.0, -0.0, -0.0, -0.0, -0.0, -0.0, -0.0, -0.0, -0.0, -0.0, -0.0, -0.0, -0.0, -0.0, -0.0, -0.0, -0.0, -0.0, -0.0, -0.0, -0.0, -0.0, -0.0, -0.0, -0.0, -0.0, -0.0, -0.0, -0.0, -0.0, -0.0, -0.0, -0.0, -0.0, -0.0, -0.0, -0.0, -0.0, -0.0, -0.0, -0.0, -0.0, -0.0, -0.0, -0.0, -0.0, -0.0, -0.0, -0.0, -0.0, -0.0, -0.0, -0.0, -0.0, -0.0, -0.0, -0.0, -0.0, -0.0, -0.0, -0.0, -0.0, -0.0, -0.0, -0.0, -0.0, -0.0, -0.0, -0.0, -0.0, -0.0, -0.0, -0.0, -0.0, -0.0, -0.0, -0.0, -0.0, -0.0, -0.0, -0.0, -0.0, 0.0, 0.0, 0.0, 0.0, 0.0, 0.0, 0.0, 0.0, 0.0, 0.0, 0.0, 0.0, 0.0, 0.0, 0.0, 0.0, 0.0, 0.0, 0.0, 0.0, 0.0, 0.0, 0.0, 0.0, 0.0, 0.0, 0.0, 0.0, 0.0, 0.0, 0.0, 0.0, 0.0, 0.0, 0.0, 0.0, 0.0, 0.0, 0.0, 0.0, 0.0, 0.0, 0.0, 0.0, 0.0, 0.0, 0.0, 0.0, 0.0, 0.0, 0.0, 0.0, 0.0, 0.0, 0.0, 0.0, 0.0, 0.0, 0.0, 0.0, 0.0, 0.0, 0.0, 0.0, 0.0, 0.0, 0.0, 0.0, 0.0, 0.0, 0.0, 0.0, 0.0, 0.0, 0.0, 0.0, 0.0, 0.0, 0.0, 0.0, 0.0, 0.0, 0.0, 0.0, 0.0, 0.0, 0.0, 0.0, 0.0, 0.0, 0.0, 0.0, 0.0, 0.0, 0.0, 0.0, 0.0, 0.0, 0.0, 0.0, 0.0, 0.0, 0.0, 0.0, 0.0, 0.0, 0.0, 0.0, 0.0, 0.0, 0.0, 0.0, 0.0, 0.0, 0.0, 0.0, 0.0, 0.0, 0.0, 0.0, 0.0, 0.0, 0.0, 0.0, -0.0, -0.0, -0.0, -0.0, -0.0, -0.0, -0.0, -0.0, -0.0, -0.0, -0.0, -0.0, -0.0, -0.0, -0.0, -0.0, -0.0, -0.0, -0.0, -0.0, -0.0, -0.0, -0.0, -0.0, -0.0, -0.0, -0.0, -0.0, -0.0, -0.0, -0.0, -0.0, -0.0, -0.0, -0.0, -0.0, -0.0, -0.0, -0.0, -0.0, -0.0, -0.0, -0.0, -0.0, -0.0, -0.0, -0.0, -0.0, -0.0, -0.0, -0.0, -0.0, -0.0, -0.0, -0.0, -0.0, -0.0, -0.0, -0.0, -0.0, -0.0, -0.0, -0.0, -0.0, -0.0, -0.0, -0.0, -0.0, -0.0, -0.0, -0.0, -0.0, -0.0, -0.0, -0.0, -0.0, -0.0, -0.0, -1.7756006070928429E-5, -1.955926027849794E-5, -2.1265642444599059E-5, -2.2878087249309936E-5, -2.4399475238503513E-5, -2.5832632877734329E-5, -2.7180332648224444E-5, -2.8445293182983732E-5, -2.9630179441154765E-5, -3.0737602918726609E-5, -3.1770121893815045E-5, -3.2730241704758869E-5, -3.3620415059333691E-5, -3.4443042373434618E-5, -3.5200472137629193E-5, -3.5895001310030509E-5, -3.652887573398812E-5, -3.7104290579141277E-5, -3.7623390804425058E-5, -3.808827164166491E-5, -3.8500979098439383E-5, -3.886351047893401E-5, -3.9177814921551905E-5, -3.9445793952087749E-5, -3.966930205131298E-5, -3.98501472358593E-5, -3.9990091651326829E-5, -4.0090852176581095E-5, -4.0154101038240283E-5, -4.0181466434390562E-5, -4.017453316660271E-5, -4.013484327935801E-5, -4.0063896706025282E-5, -3.9963151920563813E-5, -3.9834026594159355E-5, -3.9677898256031791E-5, -3.9496104957683613E-5, -3.9289945939888413E-5, -3.9060682301747689E-5, -3.8809537671172525E-5, -3.8537698876174604E-5, -3.8246316616377579E-5, 0.0, 0.0, 0.0, 0.0, 0.0, 0.0, 0.0, 0.0, 0.0, 0.0, 0.0, 0.0, 0.0, 0.0, 0.0, 0.0, 0.0, 0.0, 0.0, 0.0, 0.0, 0.0, 0.0, 0.0, 0.0, 0.0, 0.0, 0.0, 0.0, 0.0, 0.0, 0.0, 0.0, 0.0, 0.0, 0.0, 0.0, 0.0, 0.0, 0.0, 0.0, 0.0, 0.0, 0.0, 0.0, 0.0, 0.0, 0.0, 0.0, 0.0, 0.0, 0.0, 0.0, 0.0, 0.0, 0.0, 0.0, 0.0, 0.0, 0.0, 0.0, 0.0, 0.0, 0.0, 0.0, 0.0, 0.0, 0.0, 0.0, 0.0, 0.0, 0.0, 0.0, 0.0, 0.0, 0.0, 0.0, 0.0, 1.7756006070928429E-5, 1.955926027849794E-5, 2.1265642444599059E-5, 2.2878087249309936E-5, 2.4399475238503513E-5, 2.5832632877734329E-5, 2.7180332648224444E-5, 2.8445293182983732E-5, 2.9630179441154765E-5, 3.0737602918726609E-5, 3.1770121893815045E-5, 3.2730241704758869E-5, 3.3620415059333691E-5, 3.4443042373434618E-5, 3.5200472137629193E-5, 3.5895001310030509E-5, 3.652887573398812E-5, 3.7104290579141277E-5, 3.7623390804425058E-5, 3.808827164166491E-5, 3.8500979098439383E-5, 3.886351047893401E-5, 3.9177814921551905E-5, 3.9445793952087749E-5, 3.966930205131298E-5, 3.98501472358593E-5, 3.9990091651326829E-5, 4.0090852176581095E-5, 4.0154101038240283E-5, 4.0181466434390562E-5, 4.017453316660271E-5, 4.013484327935801E-5, 4.0063896706025282E-5, 3.9963151920563813E-5, 3.9834026594159355E-5, 3.9677898256031791E-5, 3.9496104957683613E-5, 3.9289945939888413E-5, 3.9060682301747689E-5, 3.8809537671172525E-5, 3.8537698876174604E-5, 3.8246316616377579E-5, 0.0, 0.0, 0.0, 0.0, -0.0, -0.0, -0.0, -0.0, -0.0, -0.0, -0.0, -0.0, -0.0, -0.0, -0.0, -0.0, -0.0, -0.0, -0.0, -0.0, -0.0, -0.0, -0.0, -0.0, -0.0, -0.0, -0.0, -0.0, -0.0, -0.0, -0.0, -0.0, -0.0, -0.0, -0.0, -0.0, -0.0, -0.0, -0.0, -0.0, -0.0, -0.0, -0.0, -0.0, -0.0, -0.0, -0.0, -0.0, -0.0, -0.0, -0.0, -0.0, -0.0, -0.0, -0.0, -0.0, -0.0, -0.0, -0.0, -0.0, -0.0, -0.0, -0.0, -0.0, -0.0, -0.0, -0.0, -0.0, -0.0, -0.0, -0.0, -0.0, -0.0, -0.0, -0.0, -0.0, -0.0, -0.0, -0.0, -0.0, -0.0, -0.0, -0.0, -0.0, -0.0, -0.0, -0.0, -0.0, -0.0, -0.0, -0.0, -0.0, -0.0, -0.0, -0.0, -0.0, -0.0, -0.0, -0.0, -0.0, -0.0, -0.0, -0.0, -0.0, -0.0, -0.0, -0.0, -0.0, -0.0, -0.0, -0.0, -0.0, -0.0, -0.0, -0.0, -0.0, -0.0, -0.0, -0.0, -0.0, -0.0, -0.0, -0.0, -0.0, 0.0, 0.0, 0.0, 0.0, 0.0, 0.0, 0.0, 0.0, 0.0, 0.0, 0.0, 0.0, 0.0, 0.0, 0.0, 0.0, 0.0, 0.0, 0.0, 0.0, 0.0, 0.0, 0.0, 0.0, 0.0, 0.0, 0.0, 0.0, 0.0, 0.0, 0.0, 0.0, 0.0, 0.0, 0.0, 0.0, 0.0, 0.0, 0.0, 0.0, 0.0, 0.0, 0.0, 0.0, 0.0, 0.0, 0.0, 0.0, 0.0, 0.0, 0.0, 0.0, 0.0, 0.0, 0.0, 0.0, 0.0, 0.0, 0.0, 0.0, 0.0, 0.0, 0.0, 0.0, 0.0, 0.0, 0.0, 0.0, 0.0, 0.0, 0.0, 0.0, 0.0, 0.0, 0.0, 0.0, 0.0, 0.0, 0.0, 0.0, 0.0, 0.0, 0.0, 0.0, 0.0, 0.0, 0.0, 0.0, 0.0, 0.0, 0.0, 0.0, 0.0, 0.0, 0.0, 0.0, 0.0, 0.0, 0.0, 0.0, 0.0, 0.0, 0.0, 0.0, 0.0, 0.0, 0.0, 0.0, 0.0, 0.0, 0.0, 0.0, 0.0, 0.0, 0.0, 0.0, 0.0, 0.0, 0.0, 0.0, 0.0, 0.0, 0.0, 0.0, -0.0, -0.0, -0.0, -0.0, -0.0, -0.0, -0.0, -0.0, -0.0, -0.0, -0.0, -0.0, -0.0, -0.0, -0.0, -0.0, -0.0, -0.0, -0.0, -0.0, -0.0, -0.0, -0.0, -0.0, -0.0, -0.0, -0.0, -0.0, -0.0, -0.0, -0.0, -0.0, -0.0, -0.0, -0.0, -0.0, -0.0, -0.0, -0.0, -0.0, -0.0, -0.0, -0.0, -0.0, -0.0, -0.0, -0.0, -0.0, -0.0, -0.0, -0.0, -0.0, -0.0, -0.0, -0.0, -0.0, -0.0, -0.0, -0.0, -0.0, -0.0, -0.0, -0.0, -0.0, -0.0, -0.0, -0.0, -0.0, -0.0, -0.0, -0.0, -0.0, -0.0, -0.0, -0.0, -0.0, -0.0, -0.0, -0.0, -1.7756006070928429E-5, -1.955926027849794E-5, -2.1265642444599059E-5, -2.2878087249309936E-5, -2.4399475238503513E-5, -2.5832632877734329E-5, -2.7180332648224444E-5, -2.8445293182983732E-5, -2.9630179441154765E-5, -3.0737602918726609E-5, -3.1770121893815045E-5, -3.2730241704758869E-5, -3.3620415059333691E-5, -3.4443042373434618E-5, -3.5200472137629193E-5, -3.5895001310030509E-5, -3.652887573398812E-5, -3.7104290579141277E-5, -3.7623390804425058E-5, -3.808827164166491E-5, -3.8500979098439383E-5, -3.886351047893401E-5, -3.9177814921551905E-5, -3.9445793952087749E-5, -3.966930205131298E-5, -3.98501472358593E-5, -3.9990091651326829E-5, -4.0090852176581095E-5, -4.0154101038240283E-5, -4.0181466434390562E-5, -4.017453316660271E-5, -4.013484327935801E-5, -4.0063896706025282E-5, -3.9963151920563813E-5, -3.9834026594159355E-5, -3.9677898256031791E-5, -3.9496104957683613E-5, -3.9289945939888413E-5, -3.9060682301747689E-5, -3.8809537671172525E-5, -3.8537698876174604E-5, 0.0, 0.0, 0.0, 0.0, 0.0, 0.0, 0.0, 0.0, 0.0, 0.0, 0.0, 0.0, 0.0, 0.0, 0.0, 0.0, 0.0, 0.0, 0.0, 0.0, 0.0, 0.0, 0.0, 0.0, 0.0, 0.0, 0.0, 0.0, 0.0, 0.0, 0.0, 0.0, 0.0, 0.0, 0.0, 0.0, 0.0, 0.0, 0.0, 0.0, 0.0, 0.0, 0.0, 0.0, 0.0, 0.0, 0.0, 0.0, 0.0, 0.0, 0.0, 0.0, 0.0, 0.0, 0.0, 0.0, 0.0, 0.0, 0.0, 0.0, 0.0, 0.0, 0.0, 0.0, 0.0, 0.0, 0.0, 0.0, 0.0, 0.0, 0.0, 0.0, 0.0, 0.0, 0.0, 0.0, 0.0, 0.0, 0.0, 1.7756006070928429E-5, 1.955926027849794E-5, 2.1265642444599059E-5, 2.2878087249309936E-5, 2.4399475238503513E-5, 2.5832632877734329E-5, 2.7180332648224444E-5, 2.8445293182983732E-5, 2.9630179441154765E-5, 3.0737602918726609E-5, 3.1770121893815045E-5, 3.2730241704758869E-5, 3.3620415059333691E-5, 3.4443042373434618E-5, 3.5200472137629193E-5, 3.5895001310030509E-5, 3.652887573398812E-5, 3.7104290579141277E-5, 3.7623390804425058E-5, 3.808827164166491E-5, 3.8500979098439383E-5, 3.886351047893401E-5, 3.9177814921551905E-5, 3.9445793952087749E-5, 3.966930205131298E-5, 3.98501472358593E-5, 3.9990091651326829E-5, 4.0090852176581095E-5, 4.0154101038240283E-5, 4.0181466434390562E-5, 4.017453316660271E-5, 4.013484327935801E-5, 4.0063896706025282E-5, 3.9963151920563813E-5, 3.9834026594159355E-5, 3.9677898256031791E-5, 3.9496104957683613E-5, 3.9289945939888413E-5, 3.9060682301747689E-5, 3.8809537671172525E-5, 3.8537698876174604E-5, 0.0, 0.0, 0.0, 0.0, -0.0, -0.0, -0.0, -0.0, -0.0, -0.0, -0.0, -0.0, -0.0, -0.0, -0.0, -0.0, -0.0, -0.0, -0.0, -0.0, -0.0, -0.0, -0.0, -0.0, -0.0, -0.0, -0.0, -0.0, -0.0, -0.0, -0.0, -0.0, -0.0, -0.0, -0.0, -0.0, -0.0, -0.0, -0.0, -0.0, -0.0, -0.0, -0.0, -0.0, -0.0, -0.0, -0.0, -0.0, -0.0, -0.0, -0.0, -0.0, -0.0, -0.0, -0.0, -0.0, -0.0, -0.0, -0.0, -0.0, -0.0, -0.0, -0.0, -0.0, -0.0, -0.0, -0.0, -0.0, -0.0, -0.0, -0.0, -0.0, -0.0, -0.0, -0.0, -0.0, -0.0, -0.0, -0.0, -0.0, -0.0, -0.0, -0.0, -0.0, -0.0, -0.0, -0.0, -0.0, -0.0, -0.0, -0.0, -0.0, -0.0, -0.0, -0.0, -0.0, -0.0, -0.0, -0.0, -0.0, -0.0, -0.0, -0.0, -0.0, -0.0, -0.0, -0.0, -0.0, -0.0, -0.0, -0.0, -0.0, -0.0, -0.0, -0.0, -0.0, -0.0, -0.0, -0.0, -0.0, -0.0, -0.0, -0.0, -0.0, 0.0, 0.0, 0.0, 0.0, 0.0, 0.0, 0.0, 0.0, 0.0, 0.0, 0.0, 0.0, 0.0, 0.0, 0.0, 0.0, 0.0, 0.0, 0.0, 0.0, 0.0, 0.0, 0.0, 0.0, 0.0, 0.0, 0.0, 0.0, 0.0, 0.0, 0.0, 0.0, 0.0, 0.0, 0.0, 0.0, 0.0, 0.0, 0.0, 0.0, 0.0, 0.0, 0.0, 0.0, 0.0, 0.0, 0.0, 0.0, 0.0, 0.0, 0.0, 0.0, 0.0, 0.0, 0.0, 0.0, 0.0, 0.0, 0.0, 0.0, 0.0, 0.0, 0.0, 0.0, 0.0, 0.0, 0.0, 0.0, 0.0, 0.0, 0.0, 0.0, 0.0, 0.0, 0.0, 0.0, 0.0, 0.0, 0.0, 0.0, 0.0, 0.0, 0.0, 0.0, 0.0, 0.0, 0.0, 0.0, 0.0, 0.0, 0.0, 0.0, 0.0, 0.0, 0.0, 0.0, 0.0, 0.0, 0.0, 0.0, 0.0, 0.0, 0.0, 0.0, 0.0, 0.0, 0.0, 0.0, 0.0, 0.0, 0.0, 0.0, 0.0, 0.0, 0.0, 0.0, 0.0, 0.0, 0.0, 0.0, 0.0, 0.0, 0.0, 0.0, -0.0, -0.0, -0.0, -0.0, -0.0, -0.0, -0.0, -0.0, -0.0, -0.0, -0.0, -0.0, -0.0, -0.0, -0.0, -0.0, -0.0, -0.0, -0.0, -0.0, -0.0, -0.0, -0.0, -0.0, -0.0, -0.0, -0.0, -0.0, -0.0, -0.0, -0.0, -0.0, -0.0, -0.0, -0.0, -0.0, -0.0, -0.0, -0.0, -0.0, -0.0, -0.0, -0.0, -0.0, -0.0, -0.0, -0.0, -0.0, -0.0, -0.0, -0.0, -0.0, -0.0, -0.0, -0.0, -0.0, -0.0, -0.0, -0.0, -0.0, -0.0, -0.0, -0.0, -0.0, -0.0, -0.0, -0.0, -0.0, -0.0, -0.0, -0.0, -0.0, -0.0, -0.0, -0.0, -0.0, -0.0, -0.0, -0.0, -0.0, -1.7756006070928429E-5, -1.955926027849794E-5, -2.1265642444599059E-5, -2.2878087249309936E-5, -2.4399475238503513E-5, -2.5832632877734329E-5, -2.7180332648224444E-5, -2.8445293182983732E-5, -2.9630179441154765E-5, -3.0737602918726609E-5, -3.1770121893815045E-5, -3.2730241704758869E-5, -3.3620415059333691E-5, -3.4443042373434618E-5, -3.5200472137629193E-5, -3.5895001310030509E-5, -3.652887573398812E-5, -3.7104290579141277E-5, -3.7623390804425058E-5, -3.808827164166491E-5, -3.8500979098439383E-5, -3.886351047893401E-5, -3.9177814921551905E-5, -3.9445793952087749E-5, -3.966930205131298E-5, -3.98501472358593E-5, -3.9990091651326829E-5, -4.0090852176581095E-5, -4.0154101038240283E-5, -4.0181466434390562E-5, -4.017453316660271E-5, -4.013484327935801E-5, -4.0063896706025282E-5, -3.9963151920563813E-5, -3.9834026594159355E-5, -3.9677898256031791E-5, -3.9496104957683613E-5, -3.9289945939888413E-5, -3.9060682301747689E-5, -3.8809537671172525E-5, 0.0, 0.0, 0.0, 0.0, 0.0, 0.0, 0.0, 0.0, 0.0, 0.0, 0.0, 0.0, 0.0, 0.0, 0.0, 0.0, 0.0, 0.0, 0.0, 0.0, 0.0, 0.0, 0.0, 0.0, 0.0, 0.0, 0.0, 0.0, 0.0, 0.0, 0.0, 0.0, 0.0, 0.0, 0.0, 0.0, 0.0, 0.0, 0.0, 0.0, 0.0, 0.0, 0.0, 0.0, 0.0, 0.0, 0.0, 0.0, 0.0, 0.0, 0.0, 0.0, 0.0, 0.0, 0.0, 0.0, 0.0, 0.0, 0.0, 0.0, 0.0, 0.0, 0.0, 0.0, 0.0, 0.0, 0.0, 0.0, 0.0, 0.0, 0.0, 0.0, 0.0, 0.0, 0.0, 0.0, 0.0, 0.0, 0.0, 0.0, 1.7756006070928429E-5, 1.955926027849794E-5, 2.1265642444599059E-5, 2.2878087249309936E-5, 2.4399475238503513E-5, 2.5832632877734329E-5, 2.7180332648224444E-5, 2.8445293182983732E-5, 2.9630179441154765E-5, 3.0737602918726609E-5, 3.1770121893815045E-5, 3.2730241704758869E-5, 3.3620415059333691E-5, 3.4443042373434618E-5, 3.5200472137629193E-5, 3.5895001310030509E-5, 3.652887573398812E-5, 3.7104290579141277E-5, 3.7623390804425058E-5, 3.808827164166491E-5, 3.8500979098439383E-5, 3.886351047893401E-5, 3.9177814921551905E-5, 3.9445793952087749E-5, 3.966930205131298E-5, 3.98501472358593E-5, 3.9990091651326829E-5, 4.0090852176581095E-5, 4.0154101038240283E-5, 4.0181466434390562E-5, 4.017453316660271E-5, 4.013484327935801E-5, 4.0063896706025282E-5, 3.9963151920563813E-5, 3.9834026594159355E-5, 3.9677898256031791E-5, 3.9496104957683613E-5, 3.9289945939888413E-5, 3.9060682301747689E-5, 3.8809537671172525E-5, 0.0, 0.0, 0.0, 0.0, -0.0, -0.0, -0.0, -0.0, -0.0, -0.0, -0.0, -0.0, -0.0, -0.0, -0.0, -0.0, -0.0, -0.0, -0.0, -0.0, -0.0, -0.0, -0.0, -0.0, -0.0, -0.0, -0.0, -0.0, -0.0, -0.0, -0.0, -0.0, -0.0, -0.0, -0.0, -0.0, -0.0, -0.0, -0.0, -0.0, -0.0, -0.0, -0.0, -0.0, -0.0, -0.0, -0.0, -0.0, -0.0, -0.0, -0.0, -0.0, -0.0, -0.0, -0.0, -0.0, -0.0, -0.0, -0.0, -0.0, -0.0, -0.0, -0.0, -0.0, -0.0, -0.0, -0.0, -0.0, -0.0, -0.0, -0.0, -0.0, -0.0, -0.0, -0.0, -0.0, -0.0, -0.0, -0.0, -0.0, -0.0, -0.0, -0.0, -0.0, -0.0, -0.0, -0.0, -0.0, -0.0, -0.0, -0.0, -0.0, -0.0, -0.0, -0.0, -0.0, -0.0, -0.0, -0.0, -0.0, -0.0, -0.0, -0.0, -0.0, -0.0, -0.0, -0.0, -0.0, -0.0, -0.0, -0.0, -0.0, -0.0, -0.0, -0.0, -0.0, -0.0, -0.0, -0.0, -0.0, -0.0, -0.0, -0.0, -0.0, 0.0, 0.0, 0.0, 0.0, 0.0, 0.0, 0.0, 0.0, 0.0, 0.0, 0.0, 0.0, 0.0, 0.0, 0.0, 0.0, 0.0, 0.0, 0.0, 0.0, 0.0, 0.0, 0.0, 0.0, 0.0, 0.0, 0.0, 0.0, 0.0, 0.0, 0.0, 0.0, 0.0, 0.0, 0.0, 0.0, 0.0, 0.0, 0.0, 0.0, 0.0, 0.0, 0.0, 0.0, 0.0, 0.0, 0.0, 0.0, 0.0, 0.0, 0.0, 0.0, 0.0, 0.0, 0.0, 0.0, 0.0, 0.0, 0.0, 0.0, 0.0, 0.0, 0.0, 0.0, 0.0, 0.0, 0.0, 0.0, 0.0, 0.0, 0.0, 0.0, 0.0, 0.0, 0.0, 0.0, 0.0, 0.0, 0.0, 0.0, 0.0, 0.0, 0.0, 0.0, 0.0, 0.0, 0.0, 0.0, 0.0, 0.0, 0.0, 0.0, 0.0, 0.0, 0.0, 0.0, 0.0, 0.0, 0.0, 0.0, 0.0, 0.0, 0.0, 0.0, 0.0, 0.0, 0.0, 0.0, 0.0, 0.0, 0.0, 0.0, 0.0, 0.0, 0.0, 0.0, 0.0, 0.0, 0.0, 0.0, 0.0, 0.0, 0.0, 0.0, -0.0, -0.0, -0.0, -0.0, -0.0, -0.0, -0.0, -0.0, -0.0, -0.0, -0.0, -0.0, -0.0, -0.0, -0.0, -0.0, -0.0, -0.0, -0.0, -0.0, -0.0, -0.0, -0.0, -0.0, -0.0, -0.0, -0.0, -0.0, -0.0, -0.0, -0.0, -0.0, -0.0, -0.0, -0.0, -0.0, -0.0, -0.0, -0.0, -0.0, -0.0, -0.0, -0.0, -0.0, -0.0, -0.0, -0.0, -0.0, -0.0, -0.0, -0.0, -0.0, -0.0, -0.0, -0.0, -0.0, -0.0, -0.0, -0.0, -0.0, -0.0, -0.0, -0.0, -0.0, -0.0, -0.0, -0.0, -0.0, -0.0, -0.0, -0.0, -0.0, -0.0, -0.0, -0.0, -0.0, -0.0, -0.0, -0.0, -0.0, -0.0, -1.7756006070928429E-5, -1.955926027849794E-5, -2.1265642444599059E-5, -2.2878087249309936E-5, -2.4399475238503513E-5, -2.5832632877734329E-5, -2.7180332648224444E-5, -2.8445293182983732E-5, -2.9630179441154765E-5, -3.0737602918726609E-5, -3.1770121893815045E-5, -3.2730241704758869E-5, -3.3620415059333691E-5, -3.4443042373434618E-5, -3.5200472137629193E-5, -3.5895001310030509E-5, -3.652887573398812E-5, -3.7104290579141277E-5, -3.7623390804425058E-5, -3.808827164166491E-5, -3.8500979098439383E-5, -3.886351047893401E-5, -3.9177814921551905E-5, -3.9445793952087749E-5, -3.966930205131298E-5, -3.98501472358593E-5, -3.9990091651326829E-5, -4.0090852176581095E-5, -4.0154101038240283E-5, -4.0181466434390562E-5, -4.017453316660271E-5, -4.013484327935801E-5, -4.0063896706025282E-5, -3.9963151920563813E-5, -3.9834026594159355E-5, -3.9677898256031791E-5, -3.9496104957683613E-5, -3.9289945939888413E-5, -3.9060682301747689E-5, 0.0, 0.0, 0.0, 0.0, 0.0, 0.0, 0.0, 0.0, 0.0, 0.0, 0.0, 0.0, 0.0, 0.0, 0.0, 0.0, 0.0, 0.0, 0.0, 0.0, 0.0, 0.0, 0.0, 0.0, 0.0, 0.0, 0.0, 0.0, 0.0, 0.0, 0.0, 0.0, 0.0, 0.0, 0.0, 0.0, 0.0, 0.0, 0.0, 0.0, 0.0, 0.0, 0.0, 0.0, 0.0, 0.0, 0.0, 0.0, 0.0, 0.0, 0.0, 0.0, 0.0, 0.0, 0.0, 0.0, 0.0, 0.0, 0.0, 0.0, 0.0, 0.0, 0.0, 0.0, 0.0, 0.0, 0.0, 0.0, 0.0, 0.0, 0.0, 0.0, 0.0, 0.0, 0.0, 0.0, 0.0, 0.0, 0.0, 0.0, 0.0, 1.7756006070928429E-5, 1.955926027849794E-5, 2.1265642444599059E-5, 2.2878087249309936E-5, 2.4399475238503513E-5, 2.5832632877734329E-5, 2.7180332648224444E-5, 2.8445293182983732E-5, 2.9630179441154765E-5, 3.0737602918726609E-5, 3.1770121893815045E-5, 3.2730241704758869E-5, 3.3620415059333691E-5, 3.4443042373434618E-5, 3.5200472137629193E-5, 3.5895001310030509E-5, 3.652887573398812E-5, 3.7104290579141277E-5, 3.7623390804425058E-5, 3.808827164166491E-5, 3.8500979098439383E-5, 3.886351047893401E-5, 3.9177814921551905E-5, 3.9445793952087749E-5, 3.966930205131298E-5, 3.98501472358593E-5, 3.9990091651326829E-5, 4.0090852176581095E-5, 4.0154101038240283E-5, 4.0181466434390562E-5, 4.017453316660271E-5, 4.013484327935801E-5, 4.0063896706025282E-5, 3.9963151920563813E-5, 3.9834026594159355E-5, 3.9677898256031791E-5, 3.9496104957683613E-5, 3.9289945939888413E-5, 3.9060682301747689E-5, 0.0, 0.0, 0.0, 0.0, -0.0, -0.0, -0.0, -0.0, -0.0, -0.0, -0.0, -0.0, -0.0, -0.0, -0.0, -0.0, -0.0, -0.0, -0.0, -0.0, -0.0, -0.0, -0.0, -0.0, -0.0, -0.0, -0.0, -0.0, -0.0, -0.0, -0.0, -0.0, -0.0, -0.0, -0.0, -0.0, -0.0, -0.0, -0.0, -0.0, -0.0, -0.0, -0.0, -0.0, -0.0, -0.0, -0.0, -0.0, -0.0, -0.0, -0.0, -0.0, -0.0, -0.0, -0.0, -0.0, -0.0, -0.0, -0.0, -0.0, -0.0, -0.0, -0.0, -0.0, -0.0, -0.0, -0.0, -0.0, -0.0, -0.0, -0.0, -0.0, -0.0, -0.0, -0.0, -0.0, -0.0, -0.0, -0.0, -0.0, -0.0, -0.0, -0.0, -0.0, -0.0, -0.0, -0.0, -0.0, -0.0, -0.0, -0.0, -0.0, -0.0, -0.0, -0.0, -0.0, -0.0, -0.0, -0.0, -0.0, -0.0, -0.0, -0.0, -0.0, -0.0, -0.0, -0.0, -0.0, -0.0, -0.0, -0.0, -0.0, -0.0, -0.0, -0.0, -0.0, -0.0, -0.0, -0.0, -0.0, -0.0, -0.0, -0.0, -0.0, 0.0, 0.0, 0.0, 0.0, 0.0, 0.0, 0.0, 0.0, 0.0, 0.0, 0.0, 0.0, 0.0, 0.0, 0.0, 0.0, 0.0, 0.0, 0.0, 0.0, 0.0, 0.0, 0.0, 0.0, 0.0, 0.0, 0.0, 0.0, 0.0, 0.0, 0.0, 0.0, 0.0, 0.0, 0.0, 0.0, 0.0, 0.0, 0.0, 0.0, 0.0, 0.0, 0.0, 0.0, 0.0, 0.0, 0.0, 0.0, 0.0, 0.0, 0.0, 0.0, 0.0, 0.0, 0.0, 0.0, 0.0, 0.0, 0.0, 0.0, 0.0, 0.0, 0.0, 0.0, 0.0, 0.0, 0.0, 0.0, 0.0, 0.0, 0.0, 0.0, 0.0, 0.0, 0.0, 0.0, 0.0, 0.0, 0.0, 0.0, 0.0, 0.0, 0.0, 0.0, 0.0, 0.0, 0.0, 0.0, 0.0, 0.0, 0.0, 0.0, 0.0, 0.0, 0.0, 0.0, 0.0, 0.0, 0.0, 0.0, 0.0, 0.0, 0.0, 0.0, 0.0, 0.0, 0.0, 0.0, 0.0, 0.0, 0.0, 0.0, 0.0, 0.0, 0.0, 0.0, 0.0, 0.0, 0.0, 0.0, 0.0, 0.0, 0.0, 0.0, -0.0, -0.0, -0.0, -0.0, -0.0, -0.0, -0.0, -0.0, -0.0, -0.0, -0.0, -0.0, -0.0, -0.0, -0.0, -0.0, -0.0, -0.0, -0.0, -0.0, -0.0, -0.0, -0.0, -0.0, -0.0, -0.0, -0.0, -0.0, -0.0, -0.0, -0.0, -0.0, -0.0, -0.0, -0.0, -0.0, -0.0, -0.0, -0.0, -0.0, -0.0, -0.0, -0.0, -0.0, -0.0, -0.0, -0.0, -0.0, -0.0, -0.0, -0.0, -0.0, -0.0, -0.0, -0.0, -0.0, -0.0, -0.0, -0.0, -0.0, -0.0, -0.0, -0.0, -0.0, -0.0, -0.0, -0.0, -0.0, -0.0, -0.0, -0.0, -0.0, -0.0, -0.0, -0.0, -0.0, -0.0, -0.0, -0.0, -0.0, -0.0, -0.0, -1.7756006070928429E-5, -1.955926027849794E-5, -2.1265642444599059E-5, -2.2878087249309936E-5, -2.4399475238503513E-5, -2.5832632877734329E-5, -2.7180332648224444E-5, -2.8445293182983732E-5, -2.9630179441154765E-5, -3.0737602918726609E-5, -3.1770121893815045E-5, -3.2730241704758869E-5, -3.3620415059333691E-5, -3.4443042373434618E-5, -3.5200472137629193E-5, -3.5895001310030509E-5, -3.652887573398812E-5, -3.7104290579141277E-5, -3.7623390804425058E-5, -3.808827164166491E-5, -3.8500979098439383E-5, -3.886351047893401E-5, -3.9177814921551905E-5, -3.9445793952087749E-5, -3.966930205131298E-5, -3.98501472358593E-5, -3.9990091651326829E-5, -4.0090852176581095E-5, -4.0154101038240283E-5, -4.0181466434390562E-5, -4.017453316660271E-5, -4.013484327935801E-5, -4.0063896706025282E-5, -3.9963151920563813E-5, -3.9834026594159355E-5, -3.9677898256031791E-5, -3.9496104957683613E-5, -3.9289945939888413E-5, 0.0, 0.0, 0.0, 0.0, 0.0, 0.0, 0.0, 0.0, 0.0, 0.0, 0.0, 0.0, 0.0, 0.0, 0.0, 0.0, 0.0, 0.0, 0.0, 0.0, 0.0, 0.0, 0.0, 0.0, 0.0, 0.0, 0.0, 0.0, 0.0, 0.0, 0.0, 0.0, 0.0, 0.0, 0.0, 0.0, 0.0, 0.0, 0.0, 0.0, 0.0, 0.0, 0.0, 0.0, 0.0, 0.0, 0.0, 0.0, 0.0, 0.0, 0.0, 0.0, 0.0, 0.0, 0.0, 0.0, 0.0, 0.0, 0.0, 0.0, 0.0, 0.0, 0.0, 0.0, 0.0, 0.0, 0.0, 0.0, 0.0, 0.0, 0.0, 0.0, 0.0, 0.0, 0.0, 0.0, 0.0, 0.0, 0.0, 0.0, 0.0, 0.0, 1.7756006070928429E-5, 1.955926027849794E-5, 2.1265642444599059E-5, 2.2878087249309936E-5, 2.4399475238503513E-5, 2.5832632877734329E-5, 2.7180332648224444E-5, 2.8445293182983732E-5, 2.9630179441154765E-5, 3.0737602918726609E-5, 3.1770121893815045E-5, 3.2730241704758869E-5, 3.3620415059333691E-5, 3.4443042373434618E-5, 3.5200472137629193E-5, 3.5895001310030509E-5, 3.652887573398812E-5, 3.7104290579141277E-5, 3.7623390804425058E-5, 3.808827164166491E-5, 3.8500979098439383E-5, 3.886351047893401E-5, 3.9177814921551905E-5, 3.9445793952087749E-5, 3.966930205131298E-5, 3.98501472358593E-5, 3.9990091651326829E-5, 4.0090852176581095E-5, 4.0154101038240283E-5, 4.0181466434390562E-5, 4.017453316660271E-5, 4.013484327935801E-5, 4.0063896706025282E-5, 3.9963151920563813E-5, 3.9834026594159355E-5, 3.9677898256031791E-5, 3.9496104957683613E-5, 3.9289945939888413E-5, 0.0, 0.0, 0.0, 0.0, -0.0, -0.0, -0.0, -0.0, -0.0, -0.0, -0.0, -0.0, -0.0, -0.0, -0.0, -0.0, -0.0, -0.0, -0.0, -0.0, -0.0, -0.0, -0.0, -0.0, -0.0, -0.0, -0.0, -0.0, -0.0, -0.0, -0.0, -0.0, -0.0, -0.0, -0.0, -0.0, -0.0, -0.0, -0.0, -0.0, -0.0, -0.0, -0.0, -0.0, -0.0, -0.0, -0.0, -0.0, -0.0, -0.0, -0.0, -0.0, -0.0, -0.0, -0.0, -0.0, -0.0, -0.0, -0.0, -0.0, -0.0, -0.0, -0.0, -0.0, -0.0, -0.0, -0.0, -0.0, -0.0, -0.0, -0.0, -0.0, -0.0, -0.0, -0.0, -0.0, -0.0, -0.0, -0.0, -0.0, -0.0, -0.0, -0.0, -0.0, -0.0, -0.0, -0.0, -0.0, -0.0, -0.0, -0.0, -0.0, -0.0, -0.0, -0.0, -0.0, -0.0, -0.0, -0.0, -0.0, -0.0, -0.0, -0.0, -0.0, -0.0, -0.0, -0.0, -0.0, -0.0, -0.0, -0.0, -0.0, -0.0, -0.0, -0.0, -0.0, -0.0, -0.0, -0.0, -0.0, -0.0, -0.0, -0.0, -0.0, 0.0, 0.0, 0.0, 0.0, 0.0, 0.0, 0.0, 0.0, 0.0, 0.0, 0.0, 0.0, 0.0, 0.0, 0.0, 0.0, 0.0, 0.0, 0.0, 0.0, 0.0, 0.0, 0.0, 0.0, 0.0, 0.0, 0.0, 0.0, 0.0, 0.0, 0.0, 0.0, 0.0, 0.0, 0.0, 0.0, 0.0, 0.0, 0.0, 0.0, 0.0, 0.0, 0.0, 0.0, 0.0, 0.0, 0.0, 0.0, 0.0, 0.0, 0.0, 0.0, 0.0, 0.0, 0.0, 0.0, 0.0, 0.0, 0.0, 0.0, 0.0, 0.0, 0.0, 0.0, 0.0, 0.0, 0.0, 0.0, 0.0, 0.0, 0.0, 0.0, 0.0, 0.0, 0.0, 0.0, 0.0, 0.0, 0.0, 0.0, 0.0, 0.0, 0.0, 0.0, 0.0, 0.0, 0.0, 0.0, 0.0, 0.0, 0.0, 0.0, 0.0, 0.0, 0.0, 0.0, 0.0, 0.0, 0.0, 0.0, 0.0, 0.0, 0.0, 0.0, 0.0, 0.0, 0.0, 0.0, 0.0, 0.0, 0.0, 0.0, 0.0, 0.0, 0.0, 0.0, 0.0, 0.0, 0.0, 0.0, 0.0, 0.0, 0.0, 0.0, -0.0, -0.0, -0.0, -0.0, -0.0, -0.0, -0.0, -0.0, -0.0, -0.0, -0.0, -0.0, -0.0, -0.0, -0.0, -0.0, -0.0, -0.0, -0.0, -0.0, -0.0, -0.0, -0.0, -0.0, -0.0, -0.0, -0.0, -0.0, -0.0, -0.0, -0.0, -0.0, -0.0, -0.0, -0.0, -0.0, -0.0, -0.0, -0.0, -0.0, -0.0, -0.0, -0.0, -0.0, -0.0, -0.0, -0.0, -0.0, -0.0, -0.0, -0.0, -0.0, -0.0, -0.0, -0.0, -0.0, -0.0, -0.0, -0.0, -0.0, -0.0, -0.0, -0.0, -0.0, -0.0, -0.0, -0.0, -0.0, -0.0, -0.0, -0.0, -0.0, -0.0, -0.0, -0.0, -0.0, -0.0, -0.0, -0.0, -0.0, -0.0, -0.0, -0.0, -1.7756006070928429E-5, -1.955926027849794E-5, -2.1265642444599059E-5, -2.2878087249309936E-5, -2.4399475238503513E-5, -2.5832632877734329E-5, -2.7180332648224444E-5, -2.8445293182983732E-5, -2.9630179441154765E-5, -3.0737602918726609E-5, -3.1770121893815045E-5, -3.2730241704758869E-5, -3.3620415059333691E-5, -3.4443042373434618E-5, -3.5200472137629193E-5, -3.5895001310030509E-5, -3.652887573398812E-5, -3.7104290579141277E-5, -3.7623390804425058E-5, -3.808827164166491E-5, -3.8500979098439383E-5, -3.886351047893401E-5, -3.9177814921551905E-5, -3.9445793952087749E-5, -3.966930205131298E-5, -3.98501472358593E-5, -3.9990091651326829E-5, -4.0090852176581095E-5, -4.0154101038240283E-5, -4.0181466434390562E-5, -4.017453316660271E-5, -4.013484327935801E-5, -4.0063896706025282E-5, -3.9963151920563813E-5, -3.9834026594159355E-5, -3.9677898256031791E-5, -3.9496104957683613E-5, 0.0, 0.0, 0.0, 0.0, 0.0, 0.0, 0.0, 0.0, 0.0, 0.0, 0.0, 0.0, 0.0, 0.0, 0.0, 0.0, 0.0, 0.0, 0.0, 0.0, 0.0, 0.0, 0.0, 0.0, 0.0, 0.0, 0.0, 0.0, 0.0, 0.0, 0.0, 0.0, 0.0, 0.0, 0.0, 0.0, 0.0, 0.0, 0.0, 0.0, 0.0, 0.0, 0.0, 0.0, 0.0, 0.0, 0.0, 0.0, 0.0, 0.0, 0.0, 0.0, 0.0, 0.0, 0.0, 0.0, 0.0, 0.0, 0.0, 0.0, 0.0, 0.0, 0.0, 0.0, 0.0, 0.0, 0.0, 0.0, 0.0, 0.0, 0.0, 0.0, 0.0, 0.0, 0.0, 0.0, 0.0, 0.0, 0.0, 0.0, 0.0, 0.0, 0.0, 1.7756006070928429E-5, 1.955926027849794E-5, 2.1265642444599059E-5, 2.2878087249309936E-5, 2.4399475238503513E-5, 2.5832632877734329E-5, 2.7180332648224444E-5, 2.8445293182983732E-5, 2.9630179441154765E-5, 3.0737602918726609E-5, 3.1770121893815045E-5, 3.2730241704758869E-5, 3.3620415059333691E-5, 3.4443042373434618E-5, 3.5200472137629193E-5, 3.5895001310030509E-5, 3.652887573398812E-5, 3.7104290579141277E-5, 3.7623390804425058E-5, 3.808827164166491E-5, 3.8500979098439383E-5, 3.886351047893401E-5, 3.9177814921551905E-5, 3.9445793952087749E-5, 3.966930205131298E-5, 3.98501472358593E-5, 3.9990091651326829E-5, 4.0090852176581095E-5, 4.0154101038240283E-5, 4.0181466434390562E-5, 4.017453316660271E-5, 4.013484327935801E-5, 4.0063896706025282E-5, 3.9963151920563813E-5, 3.9834026594159355E-5, 3.9677898256031791E-5, 3.9496104957683613E-5, 0.0, 0.0, 0.0, 0.0, -0.0, -0.0, -0.0, -0.0, -0.0, -0.0, -0.0, -0.0, -0.0, -0.0, -0.0, -0.0, -0.0, -0.0, -0.0, -0.0, -0.0, -0.0, -0.0, -0.0, -0.0, -0.0, -0.0, -0.0, -0.0, -0.0, -0.0, -0.0, -0.0, -0.0, -0.0, -0.0, -0.0, -0.0, -0.0, -0.0, -0.0, -0.0, -0.0, -0.0, -0.0, -0.0, -0.0, -0.0, -0.0, -0.0, -0.0, -0.0, -0.0, -0.0, -0.0, -0.0, -0.0, -0.0, -0.0, -0.0, -0.0, -0.0, -0.0, -0.0, -0.0, -0.0, -0.0, -0.0, -0.0, -0.0, -0.0, -0.0, -0.0, -0.0, -0.0, -0.0, -0.0, -0.0, -0.0, -0.0, -0.0, -0.0, -0.0, -0.0, -0.0, -0.0, -0.0, -0.0, -0.0, -0.0, -0.0, -0.0, -0.0, -0.0, -0.0, -0.0, -0.0, -0.0, -0.0, -0.0, -0.0, -0.0, -0.0, -0.0, -0.0, -0.0, -0.0, -0.0, -0.0, -0.0, -0.0, -0.0, -0.0, -0.0, -0.0, -0.0, -0.0, -0.0, -0.0, -0.0, -0.0, -0.0, -0.0, -0.0, 0.0, 0.0, 0.0, 0.0, 0.0, 0.0, 0.0, 0.0, 0.0, 0.0, 0.0, 0.0, 0.0, 0.0, 0.0, 0.0, 0.0, 0.0, 0.0, 0.0, 0.0, 0.0, 0.0, 0.0, 0.0, 0.0, 0.0, 0.0, 0.0, 0.0, 0.0, 0.0, 0.0, 0.0, 0.0, 0.0, 0.0, 0.0, 0.0, 0.0, 0.0, 0.0, 0.0, 0.0, 0.0, 0.0, 0.0, 0.0, 0.0, 0.0, 0.0, 0.0, 0.0, 0.0, 0.0, 0.0, 0.0, 0.0, 0.0, 0.0, 0.0, 0.0, 0.0, 0.0, 0.0, 0.0, 0.0, 0.0, 0.0, 0.0, 0.0, 0.0, 0.0, 0.0, 0.0, 0.0, 0.0, 0.0, 0.0, 0.0, 0.0, 0.0, 0.0, 0.0, 0.0, 0.0, 0.0, 0.0, 0.0, 0.0, 0.0, 0.0, 0.0, 0.0, 0.0, 0.0, 0.0, 0.0, 0.0, 0.0, 0.0, 0.0, 0.0, 0.0, 0.0, 0.0, 0.0, 0.0, 0.0, 0.0, 0.0, 0.0, 0.0, 0.0, 0.0, 0.0, 0.0, 0.0, 0.0, 0.0, 0.0, 0.0, 0.0, 0.0, -0.0, -0.0, -0.0, -0.0, -0.0, -0.0, -0.0, -0.0, -0.0, -0.0, -0.0, -0.0, -0.0, -0.0, -0.0, -0.0, -0.0, -0.0, -0.0, -0.0, -0.0, -0.0, -0.0, -0.0, -0.0, -0.0, -0.0, -0.0, -0.0, -0.0, -0.0, -0.0, -0.0, -0.0, -0.0, -0.0, -0.0, -0.0, -0.0, -0.0, -0.0, -0.0, -0.0, -0.0, -0.0, -0.0, -0.0, -0.0, -0.0, -0.0, -0.0, -0.0, -0.0, -0.0, -0.0, -0.0, -0.0, -0.0, -0.0, -0.0, -0.0, -0.0, -0.0, -0.0, -0.0, -0.0, -0.0, -0.0, -0.0, -0.0, -0.0, -0.0, -0.0, -0.0, -0.0, -0.0, -0.0, -0.0, -0.0, -0.0, -0.0, -0.0, -0.0, -0.0, -1.7756006070928429E-5, -1.955926027849794E-5, -2.1265642444599059E-5, -2.2878087249309936E-5, -2.4399475238503513E-5, -2.5832632877734329E-5, -2.7180332648224444E-5, -2.8445293182983732E-5, -2.9630179441154765E-5, -3.0737602918726609E-5, -3.1770121893815045E-5, -3.2730241704758869E-5, -3.3620415059333691E-5, -3.4443042373434618E-5, -3.5200472137629193E-5, -3.5895001310030509E-5, -3.652887573398812E-5, -3.7104290579141277E-5, -3.7623390804425058E-5, -3.808827164166491E-5, -3.8500979098439383E-5, -3.886351047893401E-5, -3.9177814921551905E-5, -3.9445793952087749E-5, -3.966930205131298E-5, -3.98501472358593E-5, -3.9990091651326829E-5, -4.0090852176581095E-5, -4.0154101038240283E-5, -4.0181466434390562E-5, -4.017453316660271E-5, -4.013484327935801E-5, -4.0063896706025282E-5, -3.9963151920563813E-5, -3.9834026594159355E-5, -3.9677898256031791E-5, 0.0, 0.0, 0.0, 0.0, 0.0, 0.0, 0.0, 0.0, 0.0, 0.0, 0.0, 0.0, 0.0, 0.0, 0.0, 0.0, 0.0, 0.0, 0.0, 0.0, 0.0, 0.0, 0.0, 0.0, 0.0, 0.0, 0.0, 0.0, 0.0, 0.0, 0.0, 0.0, 0.0, 0.0, 0.0, 0.0, 0.0, 0.0, 0.0, 0.0, 0.0, 0.0, 0.0, 0.0, 0.0, 0.0, 0.0, 0.0, 0.0, 0.0, 0.0, 0.0, 0.0, 0.0, 0.0, 0.0, 0.0, 0.0, 0.0, 0.0, 0.0, 0.0, 0.0, 0.0, 0.0, 0.0, 0.0, 0.0, 0.0, 0.0, 0.0, 0.0, 0.0, 0.0, 0.0, 0.0, 0.0, 0.0, 0.0, 0.0, 0.0, 0.0, 0.0, 0.0, 1.7756006070928429E-5, 1.955926027849794E-5, 2.1265642444599059E-5, 2.2878087249309936E-5, 2.4399475238503513E-5, 2.5832632877734329E-5, 2.7180332648224444E-5, 2.8445293182983732E-5, 2.9630179441154765E-5, 3.0737602918726609E-5, 3.1770121893815045E-5, 3.2730241704758869E-5, 3.3620415059333691E-5, 3.4443042373434618E-5, 3.5200472137629193E-5, 3.5895001310030509E-5, 3.652887573398812E-5, 3.7104290579141277E-5, 3.7623390804425058E-5, 3.808827164166491E-5, 3.8500979098439383E-5, 3.886351047893401E-5, 3.9177814921551905E-5, 3.9445793952087749E-5, 3.966930205131298E-5, 3.98501472358593E-5, 3.9990091651326829E-5, 4.0090852176581095E-5, 4.0154101038240283E-5, 4.0181466434390562E-5, 4.017453316660271E-5, 4.013484327935801E-5, 4.0063896706025282E-5, 3.9963151920563813E-5, 3.9834026594159355E-5, 3.9677898256031791E-5, 0.0, 0.0, 0.0, 0.0, -0.0, -0.0, -0.0, -0.0, -0.0, -0.0, -0.0, -0.0, -0.0, -0.0, -0.0, -0.0, -0.0, -0.0, -0.0, -0.0, -0.0, -0.0, -0.0, -0.0, -0.0, -0.0, -0.0, -0.0, -0.0, -0.0, -0.0, -0.0, -0.0, -0.0, -0.0, -0.0, -0.0, -0.0, -0.0, -0.0, -0.0, -0.0, -0.0, -0.0, -0.0, -0.0, -0.0, -0.0, -0.0, -0.0, -0.0, -0.0, -0.0, -0.0, -0.0, -0.0, -0.0, -0.0, -0.0, -0.0, -0.0, -0.0, -0.0, -0.0, -0.0, -0.0, -0.0, -0.0, -0.0, -0.0, -0.0, -0.0, -0.0, -0.0, -0.0, -0.0, -0.0, -0.0, -0.0, -0.0, -0.0, -0.0, -0.0, -0.0, -0.0, -0.0, -0.0, -0.0, -0.0, -0.0, -0.0, -0.0, -0.0, -0.0, -0.0, -0.0, -0.0, -0.0, -0.0, -0.0, -0.0, -0.0, -0.0, -0.0, -0.0, -0.0, -0.0, -0.0, -0.0, -0.0, -0.0, -0.0, -0.0, -0.0, -0.0, -0.0, -0.0, -0.0, -0.0, -0.0, -0.0, -0.0, -0.0, -0.0, 0.0, 0.0, 0.0, 0.0, 0.0, 0.0, 0.0, 0.0, 0.0, 0.0, 0.0, 0.0, 0.0, 0.0, 0.0, 0.0, 0.0, 0.0, 0.0, 0.0, 0.0, 0.0, 0.0, 0.0, 0.0, 0.0, 0.0, 0.0, 0.0, 0.0, 0.0, 0.0, 0.0, 0.0, 0.0, 0.0, 0.0, 0.0, 0.0, 0.0, 0.0, 0.0, 0.0, 0.0, 0.0, 0.0, 0.0, 0.0, 0.0, 0.0, 0.0, 0.0, 0.0, 0.0, 0.0, 0.0, 0.0, 0.0, 0.0, 0.0, 0.0, 0.0, 0.0, 0.0, 0.0, 0.0, 0.0, 0.0, 0.0, 0.0, 0.0, 0.0, 0.0, 0.0, 0.0, 0.0, 0.0, 0.0, 0.0, 0.0, 0.0, 0.0, 0.0, 0.0, 0.0, 0.0, 0.0, 0.0, 0.0, 0.0, 0.0, 0.0, 0.0, 0.0, 0.0, 0.0, 0.0, 0.0, 0.0, 0.0, 0.0, 0.0, 0.0, 0.0, 0.0, 0.0, 0.0, 0.0, 0.0, 0.0, 0.0, 0.0, 0.0, 0.0, 0.0, 0.0, 0.0, 0.0, 0.0, 0.0, 0.0, 0.0, 0.0, 0.0, -0.0, -0.0, -0.0, -0.0, -0.0, -0.0, -0.0, -0.0, -0.0, -0.0, -0.0, -0.0, -0.0, -0.0, -0.0, -0.0, -0.0, -0.0, -0.0, -0.0, -0.0, -0.0, -0.0, -0.0, -0.0, -0.0, -0.0, -0.0, -0.0, -0.0, -0.0, -0.0, -0.0, -0.0, -0.0, -0.0, -0.0, -0.0, -0.0, -0.0, -0.0, -0.0, -0.0, -0.0, -0.0, -0.0, -0.0, -0.0, -0.0, -0.0, -0.0, -0.0, -0.0, -0.0, -0.0, -0.0, -0.0, -0.0, -0.0, -0.0, -0.0, -0.0, -0.0, -0.0, -0.0, -0.0, -0.0, -0.0, -0.0, -0.0, -0.0, -0.0, -0.0, -0.0, -0.0, -0.0, -0.0, -0.0, -0.0, -0.0, -0.0, -0.0, -0.0, -0.0, -0.0, -1.7756006070928429E-5, -1.955926027849794E-5, -2.1265642444599059E-5, -2.2878087249309936E-5, -2.4399475238503513E-5, -2.5832632877734329E-5, -2.7180332648224444E-5, -2.8445293182983732E-5, -2.9630179441154765E-5, -3.0737602918726609E-5, -3.1770121893815045E-5, -3.2730241704758869E-5, -3.3620415059333691E-5, -3.4443042373434618E-5, -3.5200472137629193E-5, -3.5895001310030509E-5, -3.652887573398812E-5, -3.7104290579141277E-5, -3.7623390804425058E-5, -3.808827164166491E-5, -3.8500979098439383E-5, -3.886351047893401E-5, -3.9177814921551905E-5, -3.9445793952087749E-5, -3.966930205131298E-5, -3.98501472358593E-5, -3.9990091651326829E-5, -4.0090852176581095E-5, -4.0154101038240283E-5, -4.0181466434390562E-5, -4.017453316660271E-5, -4.013484327935801E-5, -4.0063896706025282E-5, -3.9963151920563813E-5, -3.9834026594159355E-5, 0.0, 0.0, 0.0, 0.0, 0.0, 0.0, 0.0, 0.0, 0.0, 0.0, 0.0, 0.0, 0.0, 0.0, 0.0, 0.0, 0.0, 0.0, 0.0, 0.0, 0.0, 0.0, 0.0, 0.0, 0.0, 0.0, 0.0, 0.0, 0.0, 0.0, 0.0, 0.0, 0.0, 0.0, 0.0, 0.0, 0.0, 0.0, 0.0, 0.0, 0.0, 0.0, 0.0, 0.0, 0.0, 0.0, 0.0, 0.0, 0.0, 0.0, 0.0, 0.0, 0.0, 0.0, 0.0, 0.0, 0.0, 0.0, 0.0, 0.0, 0.0, 0.0, 0.0, 0.0, 0.0, 0.0, 0.0, 0.0, 0.0, 0.0, 0.0, 0.0, 0.0, 0.0, 0.0, 0.0, 0.0, 0.0, 0.0, 0.0, 0.0, 0.0, 0.0, 0.0, 0.0, 1.7756006070928429E-5, 1.955926027849794E-5, 2.1265642444599059E-5, 2.2878087249309936E-5, 2.4399475238503513E-5, 2.5832632877734329E-5, 2.7180332648224444E-5, 2.8445293182983732E-5, 2.9630179441154765E-5, 3.0737602918726609E-5, 3.1770121893815045E-5, 3.2730241704758869E-5, 3.3620415059333691E-5, 3.4443042373434618E-5, 3.5200472137629193E-5, 3.5895001310030509E-5, 3.652887573398812E-5, 3.7104290579141277E-5, 3.7623390804425058E-5, 3.808827164166491E-5, 3.8500979098439383E-5, 3.886351047893401E-5, 3.9177814921551905E-5, 3.9445793952087749E-5, 3.966930205131298E-5, 3.98501472358593E-5, 3.9990091651326829E-5, 4.0090852176581095E-5, 4.0154101038240283E-5, 4.0181466434390562E-5, 4.017453316660271E-5, 4.013484327935801E-5, 4.0063896706025282E-5, 3.9963151920563813E-5, 3.9834026594159355E-5, 0.0, 0.0, 0.0, 0.0, -0.0, -0.0, -0.0, -0.0, -0.0, -0.0, -0.0, -0.0, -0.0, -0.0, -0.0, -0.0, -0.0, -0.0, -0.0, -0.0, -0.0, -0.0, -0.0, -0.0, -0.0, -0.0, -0.0, -0.0, -0.0, -0.0, -0.0, -0.0, -0.0, -0.0, -0.0, -0.0, -0.0, -0.0, -0.0, -0.0, -0.0, -0.0, -0.0, -0.0, -0.0, -0.0, -0.0, -0.0, -0.0, -0.0, -0.0, -0.0, -0.0, -0.0, -0.0, -0.0, -0.0, -0.0, -0.0, -0.0, -0.0, -0.0, -0.0, -0.0, -0.0, -0.0, -0.0, -0.0, -0.0, -0.0, -0.0, -0.0, -0.0, -0.0, -0.0, -0.0, -0.0, -0.0, -0.0, -0.0, -0.0, -0.0, -0.0, -0.0, -0.0, -0.0, -0.0, -0.0, -0.0, -0.0, -0.0, -0.0, -0.0, -0.0, -0.0, -0.0, -0.0, -0.0, -0.0, -0.0, -0.0, -0.0, -0.0, -0.0, -0.0, -0.0, -0.0, -0.0, -0.0, -0.0, -0.0, -0.0, -0.0, -0.0, -0.0, -0.0, -0.0, -0.0, -0.0, -0.0, -0.0, -0.0, -0.0, -0.0, 0.0, 0.0, 0.0, 0.0, 0.0, 0.0, 0.0, 0.0, 0.0, 0.0, 0.0, 0.0, 0.0, 0.0, 0.0, 0.0, 0.0, 0.0, 0.0, 0.0, 0.0, 0.0, 0.0, 0.0, 0.0, 0.0, 0.0, 0.0, 0.0, 0.0, 0.0, 0.0, 0.0, 0.0, 0.0, 0.0, 0.0, 0.0, 0.0, 0.0, 0.0, 0.0, 0.0, 0.0, 0.0, 0.0, 0.0, 0.0, 0.0, 0.0, 0.0, 0.0, 0.0, 0.0, 0.0, 0.0, 0.0, 0.0, 0.0, 0.0, 0.0, 0.0, 0.0, 0.0, 0.0, 0.0, 0.0, 0.0, 0.0, 0.0, 0.0, 0.0, 0.0, 0.0, 0.0, 0.0, 0.0, 0.0, 0.0, 0.0, 0.0, 0.0, 0.0, 0.0, 0.0, 0.0, 0.0, 0.0, 0.0, 0.0, 0.0, 0.0, 0.0, 0.0, 0.0, 0.0, 0.0, 0.0, 0.0, 0.0, 0.0, 0.0, 0.0, 0.0, 0.0, 0.0, 0.0, 0.0, 0.0, 0.0, 0.0, 0.0, 0.0, 0.0, 0.0, 0.0, 0.0, 0.0, 0.0, 0.0, 0.0, 0.0, 0.0, 0.0, -0.0, -0.0, -0.0, -0.0, -0.0, -0.0, -0.0, -0.0, -0.0, -0.0, -0.0, -0.0, -0.0, -0.0, -0.0, -0.0, -0.0, -0.0, -0.0, -0.0, -0.0, -0.0, -0.0, -0.0, -0.0, -0.0, -0.0, -0.0, -0.0, -0.0, -0.0, -0.0, -0.0, -0.0, -0.0, -0.0, -0.0, -0.0, -0.0, -0.0, -0.0, -0.0, -0.0, -0.0, -0.0, -0.0, -0.0, -0.0, -0.0, -0.0, -0.0, -0.0, -0.0, -0.0, -0.0, -0.0, -0.0, -0.0, -0.0, -0.0, -0.0, -0.0, -0.0, -0.0, -0.0, -0.0, -0.0, -0.0, -0.0, -0.0, -0.0, -0.0, -0.0, -0.0, -0.0, -0.0, -0.0, -0.0, -0.0, -0.0, -0.0, -0.0, -0.0, -0.0, -0.0, -0.0, -1.7756006070928429E-5, -1.955926027849794E-5, -2.1265642444599059E-5, -2.2878087249309936E-5, -2.4399475238503513E-5, -2.5832632877734329E-5, -2.7180332648224444E-5, -2.8445293182983732E-5, -2.9630179441154765E-5, -3.0737602918726609E-5, -3.1770121893815045E-5, -3.2730241704758869E-5, -3.3620415059333691E-5, -3.4443042373434618E-5, -3.5200472137629193E-5, -3.5895001310030509E-5, -3.652887573398812E-5, -3.7104290579141277E-5, -3.7623390804425058E-5, -3.808827164166491E-5, -3.8500979098439383E-5, -3.886351047893401E-5, -3.9177814921551905E-5, -3.9445793952087749E-5, -3.966930205131298E-5, -3.98501472358593E-5, -3.9990091651326829E-5, -4.0090852176581095E-5, -4.0154101038240283E-5, -4.0181466434390562E-5, -4.017453316660271E-5, -4.013484327935801E-5, -4.0063896706025282E-5, -3.9963151920563813E-5, 0.0, 0.0, 0.0, 0.0, 0.0, 0.0, 0.0, 0.0, 0.0, 0.0, 0.0, 0.0, 0.0, 0.0, 0.0, 0.0, 0.0, 0.0, 0.0, 0.0, 0.0, 0.0, 0.0, 0.0, 0.0, 0.0, 0.0, 0.0, 0.0, 0.0, 0.0, 0.0, 0.0, 0.0, 0.0, 0.0, 0.0, 0.0, 0.0, 0.0, 0.0, 0.0, 0.0, 0.0, 0.0, 0.0, 0.0, 0.0, 0.0, 0.0, 0.0, 0.0, 0.0, 0.0, 0.0, 0.0, 0.0, 0.0, 0.0, 0.0, 0.0, 0.0, 0.0, 0.0, 0.0, 0.0, 0.0, 0.0, 0.0, 0.0, 0.0, 0.0, 0.0, 0.0, 0.0, 0.0, 0.0, 0.0, 0.0, 0.0, 0.0, 0.0, 0.0, 0.0, 0.0, 0.0, 1.7756006070928429E-5, 1.955926027849794E-5, 2.1265642444599059E-5, 2.2878087249309936E-5, 2.4399475238503513E-5, 2.5832632877734329E-5, 2.7180332648224444E-5, 2.8445293182983732E-5, 2.9630179441154765E-5, 3.0737602918726609E-5, 3.1770121893815045E-5, 3.2730241704758869E-5, 3.3620415059333691E-5, 3.4443042373434618E-5, 3.5200472137629193E-5, 3.5895001310030509E-5, 3.652887573398812E-5, 3.7104290579141277E-5, 3.7623390804425058E-5, 3.808827164166491E-5, 3.8500979098439383E-5, 3.886351047893401E-5, 3.9177814921551905E-5, 3.9445793952087749E-5, 3.966930205131298E-5, 3.98501472358593E-5, 3.9990091651326829E-5, 4.0090852176581095E-5, 4.0154101038240283E-5, 4.0181466434390562E-5, 4.017453316660271E-5, 4.013484327935801E-5, 4.0063896706025282E-5, 3.9963151920563813E-5, 0.0, 0.0, 0.0, 0.0, -0.0, -0.0, -0.0, -0.0, -0.0, -0.0, -0.0, -0.0, -0.0, -0.0, -0.0, -0.0, -0.0, -0.0, -0.0, -0.0, -0.0, -0.0, -0.0, -0.0, -0.0, -0.0, -0.0, -0.0, -0.0, -0.0, -0.0, -0.0, -0.0, -0.0, -0.0, -0.0, -0.0, -0.0, -0.0, -0.0, -0.0, -0.0, -0.0, -0.0, -0.0, -0.0, -0.0, -0.0, -0.0, -0.0, -0.0, -0.0, -0.0, -0.0, -0.0, -0.0, -0.0, -0.0, -0.0, -0.0, -0.0, -0.0, -0.0, -0.0, -0.0, -0.0, -0.0, -0.0, -0.0, -0.0, -0.0, -0.0, -0.0, -0.0, -0.0, -0.0, -0.0, -0.0, -0.0, -0.0, -0.0, -0.0, -0.0, -0.0, -0.0, -0.0, -0.0, -0.0, -0.0, -0.0, -0.0, -0.0, -0.0, -0.0, -0.0, -0.0, -0.0, -0.0, -0.0, -0.0, -0.0, -0.0, -0.0, -0.0, -0.0, -0.0, -0.0, -0.0, -0.0, -0.0, -0.0, -0.0, -0.0, -0.0, -0.0, -0.0, -0.0, -0.0, -0.0, -0.0, -0.0, -0.0, -0.0, -0.0, 0.0, 0.0, 0.0, 0.0, 0.0, 0.0, 0.0, 0.0, 0.0, 0.0, 0.0, 0.0, 0.0, 0.0, 0.0, 0.0, 0.0, 0.0, 0.0, 0.0, 0.0, 0.0, 0.0, 0.0, 0.0, 0.0, 0.0, 0.0, 0.0, 0.0, 0.0, 0.0, 0.0, 0.0, 0.0, 0.0, 0.0, 0.0, 0.0, 0.0, 0.0, 0.0, 0.0, 0.0, 0.0, 0.0, 0.0, 0.0, 0.0, 0.0, 0.0, 0.0, 0.0, 0.0, 0.0, 0.0, 0.0, 0.0, 0.0, 0.0, 0.0, 0.0, 0.0, 0.0, 0.0, 0.0, 0.0, 0.0, 0.0, 0.0, 0.0, 0.0, 0.0, 0.0, 0.0, 0.0, 0.0, 0.0, 0.0, 0.0, 0.0, 0.0, 0.0, 0.0, 0.0, 0.0, 0.0, 0.0, 0.0, 0.0, 0.0, 0.0, 0.0, 0.0, 0.0, 0.0, 0.0, 0.0, 0.0, 0.0, 0.0, 0.0, 0.0, 0.0, 0.0, 0.0, 0.0, 0.0, 0.0, 0.0, 0.0, 0.0, 0.0, 0.0, 0.0, 0.0, 0.0, 0.0, 0.0, 0.0, 0.0, 0.0, 0.0, 0.0, -0.0, -0.0, -0.0, -0.0, -0.0, -0.0, -0.0, -0.0, -0.0, -0.0, -0.0, -0.0, -0.0, -0.0, -0.0, -0.0, -0.0, -0.0, -0.0, -0.0, -0.0, -0.0, -0.0, -0.0, -0.0, -0.0, -0.0, -0.0, -0.0, -0.0, -0.0, -0.0, -0.0, -0.0, -0.0, -0.0, -0.0, -0.0, -0.0, -0.0, -0.0, -0.0, -0.0, -0.0, -0.0, -0.0, -0.0, -0.0, -0.0, -0.0, -0.0, -0.0, -0.0, -0.0, -0.0, -0.0, -0.0, -0.0, -0.0, -0.0, -0.0, -0.0, -0.0, -0.0, -0.0, -0.0, -0.0, -0.0, -0.0, -0.0, -0.0, -0.0, -0.0, -0.0, -0.0, -0.0, -0.0, -0.0, -0.0, -0.0, -0.0, -0.0, -0.0, -0.0, -0.0, -0.0, -0.0, -1.7756006070928429E-5, -1.955926027849794E-5, -2.1265642444599059E-5, -2.2878087249309936E-5, -2.4399475238503513E-5, -2.5832632877734329E-5, -2.7180332648224444E-5, -2.8445293182983732E-5, -2.9630179441154765E-5, -3.0737602918726609E-5, -3.1770121893815045E-5, -3.2730241704758869E-5, -3.3620415059333691E-5, -3.4443042373434618E-5, -3.5200472137629193E-5, -3.5895001310030509E-5, -3.652887573398812E-5, -3.7104290579141277E-5, -3.7623390804425058E-5, -3.808827164166491E-5, -3.8500979098439383E-5, -3.886351047893401E-5, -3.9177814921551905E-5, -3.9445793952087749E-5, -3.966930205131298E-5, -3.98501472358593E-5, -3.9990091651326829E-5, -4.0090852176581095E-5, -4.0154101038240283E-5, -4.0181466434390562E-5, -4.017453316660271E-5, -4.013484327935801E-5, -4.0063896706025282E-5, 0.0, 0.0, 0.0, 0.0, 0.0, 0.0, 0.0, 0.0, 0.0, 0.0, 0.0, 0.0, 0.0, 0.0, 0.0, 0.0, 0.0, 0.0, 0.0, 0.0, 0.0, 0.0, 0.0, 0.0, 0.0, 0.0, 0.0, 0.0, 0.0, 0.0, 0.0, 0.0, 0.0, 0.0, 0.0, 0.0, 0.0, 0.0, 0.0, 0.0, 0.0, 0.0, 0.0, 0.0, 0.0, 0.0, 0.0, 0.0, 0.0, 0.0, 0.0, 0.0, 0.0, 0.0, 0.0, 0.0, 0.0, 0.0, 0.0, 0.0, 0.0, 0.0, 0.0, 0.0, 0.0, 0.0, 0.0, 0.0, 0.0, 0.0, 0.0, 0.0, 0.0, 0.0, 0.0, 0.0, 0.0, 0.0, 0.0, 0.0, 0.0, 0.0, 0.0, 0.0, 0.0, 0.0, 0.0, 1.7756006070928429E-5, 1.955926027849794E-5, 2.1265642444599059E-5, 2.2878087249309936E-5, 2.4399475238503513E-5, 2.5832632877734329E-5, 2.7180332648224444E-5, 2.8445293182983732E-5, 2.9630179441154765E-5, 3.0737602918726609E-5, 3.1770121893815045E-5, 3.2730241704758869E-5, 3.3620415059333691E-5, 3.4443042373434618E-5, 3.5200472137629193E-5, 3.5895001310030509E-5, 3.652887573398812E-5, 3.7104290579141277E-5, 3.7623390804425058E-5, 3.808827164166491E-5, 3.8500979098439383E-5, 3.886351047893401E-5, 3.9177814921551905E-5, 3.9445793952087749E-5, 3.966930205131298E-5, 3.98501472358593E-5, 3.9990091651326829E-5, 4.0090852176581095E-5, 4.0154101038240283E-5, 4.0181466434390562E-5, 4.017453316660271E-5, 4.013484327935801E-5, 4.0063896706025282E-5, 0.0, 0.0, 0.0, 0.0, -0.0, -0.0, -0.0, -0.0, -0.0, -0.0, -0.0, -0.0, -0.0, -0.0, -0.0, -0.0, -0.0, -0.0, -0.0, -0.0, -0.0, -0.0, -0.0, -0.0, -0.0, -0.0, -0.0, -0.0, -0.0, -0.0, -0.0, -0.0, -0.0, -0.0, -0.0, -0.0, -0.0, -0.0, -0.0, -0.0, -0.0, -0.0, -0.0, -0.0, -0.0, -0.0, -0.0, -0.0, -0.0, -0.0, -0.0, -0.0, -0.0, -0.0, -0.0, -0.0, -0.0, -0.0, -0.0, -0.0, -0.0, -0.0, -0.0, -0.0, -0.0, -0.0, -0.0, -0.0, -0.0, -0.0, -0.0, -0.0, -0.0, -0.0, -0.0, -0.0, -0.0, -0.0, -0.0, -0.0, -0.0, -0.0, -0.0, -0.0, -0.0, -0.0, -0.0, -0.0, -0.0, -0.0, -0.0, -0.0, -0.0, -0.0, -0.0, -0.0, -0.0, -0.0, -0.0, -0.0, -0.0, -0.0, -0.0, -0.0, -0.0, -0.0, -0.0, -0.0, -0.0, -0.0, -0.0, -0.0, -0.0, -0.0, -0.0, -0.0, -0.0, -0.0, -0.0, -0.0, -0.0, -0.0, -0.0, -0.0, 0.0, 0.0, 0.0, 0.0, 0.0, 0.0, 0.0, 0.0, 0.0, 0.0, 0.0, 0.0, 0.0, 0.0, 0.0, 0.0, 0.0, 0.0, 0.0, 0.0, 0.0, 0.0, 0.0, 0.0, 0.0, 0.0, 0.0, 0.0, 0.0, 0.0, 0.0, 0.0, 0.0, 0.0, 0.0, 0.0, 0.0, 0.0, 0.0, 0.0, 0.0, 0.0, 0.0, 0.0, 0.0, 0.0, 0.0, 0.0, 0.0, 0.0, 0.0, 0.0, 0.0, 0.0, 0.0, 0.0, 0.0, 0.0, 0.0, 0.0, 0.0, 0.0, 0.0, 0.0, 0.0, 0.0, 0.0, 0.0, 0.0, 0.0, 0.0, 0.0, 0.0, 0.0, 0.0, 0.0, 0.0, 0.0, 0.0, 0.0, 0.0, 0.0, 0.0, 0.0, 0.0, 0.0, 0.0, 0.0, 0.0, 0.0, 0.0, 0.0, 0.0, 0.0, 0.0, 0.0, 0.0, 0.0, 0.0, 0.0, 0.0, 0.0, 0.0, 0.0, 0.0, 0.0, 0.0, 0.0, 0.0, 0.0, 0.0, 0.0, 0.0, 0.0, 0.0, 0.0, 0.0, 0.0, 0.0, 0.0, 0.0, 0.0, 0.0, 0.0, -0.0, -0.0, -0.0, -0.0, -0.0, -0.0, -0.0, -0.0, -0.0, -0.0, -0.0, -0.0, -0.0, -0.0, -0.0, -0.0, -0.0, -0.0, -0.0, -0.0, -0.0, -0.0, -0.0, -0.0, -0.0, -0.0, -0.0, -0.0, -0.0, -0.0, -0.0, -0.0, -0.0, -0.0, -0.0, -0.0, -0.0, -0.0, -0.0, -0.0, -0.0, -0.0, -0.0, -0.0, -0.0, -0.0, -0.0, -0.0, -0.0, -0.0, -0.0, -0.0, -0.0, -0.0, -0.0, -0.0, -0.0, -0.0, -0.0, -0.0, -0.0, -0.0, -0.0, -0.0, -0.0, -0.0, -0.0, -0.0, -0.0, -0.0, -0.0, -0.0, -0.0, -0.0, -0.0, -0.0, -0.0, -0.0, -0.0, -0.0, -0.0, -0.0, -0.0, -0.0, -0.0, -0.0, -0.0, -0.0, -1.7756006070928429E-5, -1.955926027849794E-5, -2.1265642444599059E-5, -2.2878087249309936E-5, -2.4399475238503513E-5, -2.5832632877734329E-5, -2.7180332648224444E-5, -2.8445293182983732E-5, -2.9630179441154765E-5, -3.0737602918726609E-5, -3.1770121893815045E-5, -3.2730241704758869E-5, -3.3620415059333691E-5, -3.4443042373434618E-5, -3.5200472137629193E-5, -3.5895001310030509E-5, -3.652887573398812E-5, -3.7104290579141277E-5, -3.7623390804425058E-5, -3.808827164166491E-5, -3.8500979098439383E-5, -3.886351047893401E-5, -3.9177814921551905E-5, -3.9445793952087749E-5, -3.966930205131298E-5, -3.98501472358593E-5, -3.9990091651326829E-5, -4.0090852176581095E-5, -4.0154101038240283E-5, -4.0181466434390562E-5, -4.017453316660271E-5, -4.013484327935801E-5, 0.0, 0.0, 0.0, 0.0, 0.0, 0.0, 0.0, 0.0, 0.0, 0.0, 0.0, 0.0, 0.0, 0.0, 0.0, 0.0, 0.0, 0.0, 0.0, 0.0, 0.0, 0.0, 0.0, 0.0, 0.0, 0.0, 0.0, 0.0, 0.0, 0.0, 0.0, 0.0, 0.0, 0.0, 0.0, 0.0, 0.0, 0.0, 0.0, 0.0, 0.0, 0.0, 0.0, 0.0, 0.0, 0.0, 0.0, 0.0, 0.0, 0.0, 0.0, 0.0, 0.0, 0.0, 0.0, 0.0, 0.0, 0.0, 0.0, 0.0, 0.0, 0.0, 0.0, 0.0, 0.0, 0.0, 0.0, 0.0, 0.0, 0.0, 0.0, 0.0, 0.0, 0.0, 0.0, 0.0, 0.0, 0.0, 0.0, 0.0, 0.0, 0.0, 0.0, 0.0, 0.0, 0.0, 0.0, 0.0, 1.7756006070928429E-5, 1.955926027849794E-5, 2.1265642444599059E-5, 2.2878087249309936E-5, 2.4399475238503513E-5, 2.5832632877734329E-5, 2.7180332648224444E-5, 2.8445293182983732E-5, 2.9630179441154765E-5, 3.0737602918726609E-5, 3.1770121893815045E-5, 3.2730241704758869E-5, 3.3620415059333691E-5, 3.4443042373434618E-5, 3.5200472137629193E-5, 3.5895001310030509E-5, 3.652887573398812E-5, 3.7104290579141277E-5, 3.7623390804425058E-5, 3.808827164166491E-5, 3.8500979098439383E-5, 3.886351047893401E-5, 3.9177814921551905E-5, 3.9445793952087749E-5, 3.966930205131298E-5, 3.98501472358593E-5, 3.9990091651326829E-5, 4.0090852176581095E-5, 4.0154101038240283E-5, 4.0181466434390562E-5, 4.017453316660271E-5, 4.013484327935801E-5, 0.0, 0.0, 0.0, 0.0, -0.0, -0.0, -0.0, -0.0, -0.0, -0.0, -0.0, -0.0, -0.0, -0.0, -0.0, -0.0, -0.0, -0.0, -0.0, -0.0, -0.0, -0.0, -0.0, -0.0, -0.0, -0.0, -0.0, -0.0, -0.0, -0.0, -0.0, -0.0, -0.0, -0.0, -0.0, -0.0, -0.0, -0.0, -0.0, -0.0, -0.0, -0.0, -0.0, -0.0, -0.0, -0.0, -0.0, -0.0, -0.0, -0.0, -0.0, -0.0, -0.0, -0.0, -0.0, -0.0, -0.0, -0.0, -0.0, -0.0, -0.0, -0.0, -0.0, -0.0, -0.0, -0.0, -0.0, -0.0, -0.0, -0.0, -0.0, -0.0, -0.0, -0.0, -0.0, -0.0, -0.0, -0.0, -0.0, -0.0, -0.0, -0.0, -0.0, -0.0, -0.0, -0.0, -0.0, -0.0, -0.0, -0.0, -0.0, -0.0, -0.0, -0.0, -0.0, -0.0, -0.0, -0.0, -0.0, -0.0, -0.0, -0.0, -0.0, -0.0, -0.0, -0.0, -0.0, -0.0, -0.0, -0.0, -0.0, -0.0, -0.0, -0.0, -0.0, -0.0, -0.0, -0.0, -0.0, -0.0, -0.0, -0.0, -0.0, -0.0, 0.0, 0.0, 0.0, 0.0, 0.0, 0.0, 0.0, 0.0, 0.0, 0.0, 0.0, 0.0, 0.0, 0.0, 0.0, 0.0, 0.0, 0.0, 0.0, 0.0, 0.0, 0.0, 0.0, 0.0, 0.0, 0.0, 0.0, 0.0, 0.0, 0.0, 0.0, 0.0, 0.0, 0.0, 0.0, 0.0, 0.0, 0.0, 0.0, 0.0, 0.0, 0.0, 0.0, 0.0, 0.0, 0.0, 0.0, 0.0, 0.0, 0.0, 0.0, 0.0, 0.0, 0.0, 0.0, 0.0, 0.0, 0.0, 0.0, 0.0, 0.0, 0.0, 0.0, 0.0, 0.0, 0.0, 0.0, 0.0, 0.0, 0.0, 0.0, 0.0, 0.0, 0.0, 0.0, 0.0, 0.0, 0.0, 0.0, 0.0, 0.0, 0.0, 0.0, 0.0, 0.0, 0.0, 0.0, 0.0, 0.0, 0.0, 0.0, 0.0, 0.0, 0.0, 0.0, 0.0, 0.0, 0.0, 0.0, 0.0, 0.0, 0.0, 0.0, 0.0, 0.0, 0.0, 0.0, 0.0, 0.0, 0.0, 0.0, 0.0, 0.0, 0.0, 0.0, 0.0, 0.0, 0.0, 0.0, 0.0, 0.0, 0.0, 0.0, 0.0, -0.0, -0.0, -0.0, -0.0, -0.0, -0.0, -0.0, -0.0, -0.0, -0.0, -0.0, -0.0, -0.0, -0.0, -0.0, -0.0, -0.0, -0.0, -0.0, -0.0, -0.0, -0.0, -0.0, -0.0, -0.0, -0.0, -0.0, -0.0, -0.0, -0.0, -0.0, -0.0, -0.0, -0.0, -0.0, -0.0, -0.0, -0.0, -0.0, -0.0, -0.0, -0.0, -0.0, -0.0, -0.0, -0.0, -0.0, -0.0, -0.0, -0.0, -0.0, -0.0, -0.0, -0.0, -0.0, -0.0, -0.0, -0.0, -0.0, -0.0, -0.0, -0.0, -0.0, -0.0, -0.0, -0.0, -0.0, -0.0, -0.0, -0.0, -0.0, -0.0, -0.0, -0.0, -0.0, -0.0, -0.0, -0.0, -0.0, -0.0, -0.0, -0.0, -0.0, -0.0, -0.0, -0.0, -0.0, -0.0, -0.0, -1.7756006070928429E-5, -1.955926027849794E-5, -2.1265642444599059E-5, -2.2878087249309936E-5, -2.4399475238503513E-5, -2.5832632877734329E-5, -2.7180332648224444E-5, -2.8445293182983732E-5, -2.9630179441154765E-5, -3.0737602918726609E-5, -3.1770121893815045E-5, -3.2730241704758869E-5, -3.3620415059333691E-5, -3.4443042373434618E-5, -3.5200472137629193E-5, -3.5895001310030509E-5, -3.652887573398812E-5, -3.7104290579141277E-5, -3.7623390804425058E-5, -3.808827164166491E-5, -3.8500979098439383E-5, -3.886351047893401E-5, -3.9177814921551905E-5, -3.9445793952087749E-5, -3.966930205131298E-5, -3.98501472358593E-5, -3.9990091651326829E-5, -4.0090852176581095E-5, -4.0154101038240283E-5, -4.0181466434390562E-5, -4.017453316660271E-5, 0.0, 0.0, 0.0, 0.0, 0.0, 0.0, 0.0, 0.0, 0.0, 0.0, 0.0, 0.0, 0.0, 0.0, 0.0, 0.0, 0.0, 0.0, 0.0, 0.0, 0.0, 0.0, 0.0, 0.0, 0.0, 0.0, 0.0, 0.0, 0.0, 0.0, 0.0, 0.0, 0.0, 0.0, 0.0, 0.0, 0.0, 0.0, 0.0, 0.0, 0.0, 0.0, 0.0, 0.0, 0.0, 0.0, 0.0, 0.0, 0.0, 0.0, 0.0, 0.0, 0.0, 0.0, 0.0, 0.0, 0.0, 0.0, 0.0, 0.0, 0.0, 0.0, 0.0, 0.0, 0.0, 0.0, 0.0, 0.0, 0.0, 0.0, 0.0, 0.0, 0.0, 0.0, 0.0, 0.0, 0.0, 0.0, 0.0, 0.0, 0.0, 0.0, 0.0, 0.0, 0.0, 0.0, 0.0, 0.0, 0.0, 1.7756006070928429E-5, 1.955926027849794E-5, 2.1265642444599059E-5, 2.2878087249309936E-5, 2.4399475238503513E-5, 2.5832632877734329E-5, 2.7180332648224444E-5, 2.8445293182983732E-5, 2.9630179441154765E-5, 3.0737602918726609E-5, 3.1770121893815045E-5, 3.2730241704758869E-5, 3.3620415059333691E-5, 3.4443042373434618E-5, 3.5200472137629193E-5, 3.5895001310030509E-5, 3.652887573398812E-5, 3.7104290579141277E-5, 3.7623390804425058E-5, 3.808827164166491E-5, 3.8500979098439383E-5, 3.886351047893401E-5, 3.9177814921551905E-5, 3.9445793952087749E-5, 3.966930205131298E-5, 3.98501472358593E-5, 3.9990091651326829E-5, 4.0090852176581095E-5, 4.0154101038240283E-5, 4.0181466434390562E-5, 4.017453316660271E-5, 0.0, 0.0, 0.0, 0.0, -0.0, -0.0, -0.0, -0.0, -0.0, -0.0, -0.0, -0.0, -0.0, -0.0, -0.0, -0.0, -0.0, -0.0, -0.0, -0.0, -0.0, -0.0, -0.0, -0.0, -0.0, -0.0, -0.0, -0.0, -0.0, -0.0, -0.0, -0.0, -0.0, -0.0, -0.0, -0.0, -0.0, -0.0, -0.0, -0.0, -0.0, -0.0, -0.0, -0.0, -0.0, -0.0, -0.0, -0.0, -0.0, -0.0, -0.0, -0.0, -0.0, -0.0, -0.0, -0.0, -0.0, -0.0, -0.0, -0.0, -0.0, -0.0, -0.0, -0.0, -0.0, -0.0, -0.0, -0.0, -0.0, -0.0, -0.0, -0.0, -0.0, -0.0, -0.0, -0.0, -0.0, -0.0, -0.0, -0.0, -0.0, -0.0, -0.0, -0.0, -0.0, -0.0, -0.0, -0.0, -0.0, -0.0, -0.0, -0.0, -0.0, -0.0, -0.0, -0.0, -0.0, -0.0, -0.0, -0.0, -0.0, -0.0, -0.0, -0.0, -0.0, -0.0, -0.0, -0.0, -0.0, -0.0, -0.0, -0.0, -0.0, -0.0, -0.0, -0.0, -0.0, -0.0, -0.0, -0.0, -0.0, -0.0, -0.0, -0.0, 0.0, 0.0, 0.0, 0.0, 0.0, 0.0, 0.0, 0.0, 0.0, 0.0, 0.0, 0.0, 0.0, 0.0, 0.0, 0.0, 0.0, 0.0, 0.0, 0.0, 0.0, 0.0, 0.0, 0.0, 0.0, 0.0, 0.0, 0.0, 0.0, 0.0, 0.0, 0.0, 0.0, 0.0, 0.0, 0.0, 0.0, 0.0, 0.0, 0.0, 0.0, 0.0, 0.0, 0.0, 0.0, 0.0, 0.0, 0.0, 0.0, 0.0, 0.0, 0.0, 0.0, 0.0, 0.0, 0.0, 0.0, 0.0, 0.0, 0.0, 0.0, 0.0, 0.0, 0.0, 0.0, 0.0, 0.0, 0.0, 0.0, 0.0, 0.0, 0.0, 0.0, 0.0, 0.0, 0.0, 0.0, 0.0, 0.0, 0.0, 0.0, 0.0, 0.0, 0.0, 0.0, 0.0, 0.0, 0.0, 0.0, 0.0, 0.0, 0.0, 0.0, 0.0, 0.0, 0.0, 0.0, 0.0, 0.0, 0.0, 0.0, 0.0, 0.0, 0.0, 0.0, 0.0, 0.0, 0.0, 0.0, 0.0, 0.0, 0.0, 0.0, 0.0, 0.0, 0.0, 0.0, 0.0, 0.0, 0.0, 0.0, 0.0, 0.0, 0.0, -0.0, -0.0, -0.0, -0.0, -0.0, -0.0, -0.0, -0.0, -0.0, -0.0, -0.0, -0.0, -0.0, -0.0, -0.0, -0.0, -0.0, -0.0, -0.0, -0.0, -0.0, -0.0, -0.0, -0.0, -0.0, -0.0, -0.0, -0.0, -0.0, -0.0, -0.0, -0.0, -0.0, -0.0, -0.0, -0.0, -0.0, -0.0, -0.0, -0.0, -0.0, -0.0, -0.0, -0.0, -0.0, -0.0, -0.0, -0.0, -0.0, -0.0, -0.0, -0.0, -0.0, -0.0, -0.0, -0.0, -0.0, -0.0, -0.0, -0.0, -0.0, -0.0, -0.0, -0.0, -0.0, -0.0, -0.0, -0.0, -0.0, -0.0, -0.0, -0.0, -0.0, -0.0, -0.0, -0.0, -0.0, -0.0, -0.0, -0.0, -0.0, -0.0, -0.0, -0.0, -0.0, -0.0, -0.0, -0.0, -0.0, -0.0, -1.7756006070928429E-5, -1.955926027849794E-5, -2.1265642444599059E-5, -2.2878087249309936E-5, -2.4399475238503513E-5, -2.5832632877734329E-5, -2.7180332648224444E-5, -2.8445293182983732E-5, -2.9630179441154765E-5, -3.0737602918726609E-5, -3.1770121893815045E-5, -3.2730241704758869E-5, -3.3620415059333691E-5, -3.4443042373434618E-5, -3.5200472137629193E-5, -3.5895001310030509E-5, -3.652887573398812E-5, -3.7104290579141277E-5, -3.7623390804425058E-5, -3.808827164166491E-5, -3.8500979098439383E-5, -3.886351047893401E-5, -3.9177814921551905E-5, -3.9445793952087749E-5, -3.966930205131298E-5, -3.98501472358593E-5, -3.9990091651326829E-5, -4.0090852176581095E-5, -4.0154101038240283E-5, -4.0181466434390562E-5, 0.0, 0.0, 0.0, 0.0, 0.0, 0.0, 0.0, 0.0, 0.0, 0.0, 0.0, 0.0, 0.0, 0.0, 0.0, 0.0, 0.0, 0.0, 0.0, 0.0, 0.0, 0.0, 0.0, 0.0, 0.0, 0.0, 0.0, 0.0, 0.0, 0.0, 0.0, 0.0, 0.0, 0.0, 0.0, 0.0, 0.0, 0.0, 0.0, 0.0, 0.0, 0.0, 0.0, 0.0, 0.0, 0.0, 0.0, 0.0, 0.0, 0.0, 0.0, 0.0, 0.0, 0.0, 0.0, 0.0, 0.0, 0.0, 0.0, 0.0, 0.0, 0.0, 0.0, 0.0, 0.0, 0.0, 0.0, 0.0, 0.0, 0.0, 0.0, 0.0, 0.0, 0.0, 0.0, 0.0, 0.0, 0.0, 0.0, 0.0, 0.0, 0.0, 0.0, 0.0, 0.0, 0.0, 0.0, 0.0, 0.0, 0.0, 1.7756006070928429E-5, 1.955926027849794E-5, 2.1265642444599059E-5, 2.2878087249309936E-5, 2.4399475238503513E-5, 2.5832632877734329E-5, 2.7180332648224444E-5, 2.8445293182983732E-5, 2.9630179441154765E-5, 3.0737602918726609E-5, 3.1770121893815045E-5, 3.2730241704758869E-5, 3.3620415059333691E-5, 3.4443042373434618E-5, 3.5200472137629193E-5, 3.5895001310030509E-5, 3.652887573398812E-5, 3.7104290579141277E-5, 3.7623390804425058E-5, 3.808827164166491E-5, 3.8500979098439383E-5, 3.886351047893401E-5, 3.9177814921551905E-5, 3.9445793952087749E-5, 3.966930205131298E-5, 3.98501472358593E-5, 3.9990091651326829E-5, 4.0090852176581095E-5, 4.0154101038240283E-5, 4.0181466434390562E-5, 0.0, 0.0, 0.0, 0.0, -0.0, -0.0, -0.0, -0.0, -0.0, -0.0, -0.0, -0.0, -0.0, -0.0, -0.0, -0.0, -0.0, -0.0, -0.0, -0.0, -0.0, -0.0, -0.0, -0.0, -0.0, -0.0, -0.0, -0.0, -0.0, -0.0, -0.0, -0.0, -0.0, -0.0, -0.0, -0.0, -0.0, -0.0, -0.0, -0.0, -0.0, -0.0, -0.0, -0.0, -0.0, -0.0, -0.0, -0.0, -0.0, -0.0, -0.0, -0.0, -0.0, -0.0, -0.0, -0.0, -0.0, -0.0, -0.0, -0.0, -0.0, -0.0, -0.0, -0.0, -0.0, -0.0, -0.0, -0.0, -0.0, -0.0, -0.0, -0.0, -0.0, -0.0, -0.0, -0.0, -0.0, -0.0, -0.0, -0.0, -0.0, -0.0, -0.0, -0.0, -0.0, -0.0, -0.0, -0.0, -0.0, -0.0, -0.0, -0.0, -0.0, -0.0, -0.0, -0.0, -0.0, -0.0, -0.0, -0.0, -0.0, -0.0, -0.0, -0.0, -0.0, -0.0, -0.0, -0.0, -0.0, -0.0, -0.0, -0.0, -0.0, -0.0, -0.0, -0.0, -0.0, -0.0, -0.0, -0.0, -0.0, -0.0, -0.0, -0.0, 0.0, 0.0, 0.0, 0.0, 0.0, 0.0, 0.0, 0.0, 0.0, 0.0, 0.0, 0.0, 0.0, 0.0, 0.0, 0.0, 0.0, 0.0, 0.0, 0.0, 0.0, 0.0, 0.0, 0.0, 0.0, 0.0, 0.0, 0.0, 0.0, 0.0, 0.0, 0.0, 0.0, 0.0, 0.0, 0.0, 0.0, 0.0, 0.0, 0.0, 0.0, 0.0, 0.0, 0.0, 0.0, 0.0, 0.0, 0.0, 0.0, 0.0, 0.0, 0.0, 0.0, 0.0, 0.0, 0.0, 0.0, 0.0, 0.0, 0.0, 0.0, 0.0, 0.0, 0.0, 0.0, 0.0, 0.0, 0.0, 0.0, 0.0, 0.0, 0.0, 0.0, 0.0, 0.0, 0.0, 0.0, 0.0, 0.0, 0.0, 0.0, 0.0, 0.0, 0.0, 0.0, 0.0, 0.0, 0.0, 0.0, 0.0, 0.0, 0.0, 0.0, 0.0, 0.0, 0.0, 0.0, 0.0, 0.0, 0.0, 0.0, 0.0, 0.0, 0.0, 0.0, 0.0, 0.0, 0.0, 0.0, 0.0, 0.0, 0.0, 0.0, 0.0, 0.0, 0.0, 0.0, 0.0, 0.0, 0.0, 0.0, 0.0, 0.0, 0.0, -0.0, -0.0, -0.0, -0.0, -0.0, -0.0, -0.0, -0.0, -0.0, -0.0, -0.0, -0.0, -0.0, -0.0, -0.0, -0.0, -0.0, -0.0, -0.0, -0.0, -0.0, -0.0, -0.0, -0.0, -0.0, -0.0, -0.0, -0.0, -0.0, -0.0, -0.0, -0.0, -0.0, -0.0, -0.0, -0.0, -0.0, -0.0, -0.0, -0.0, -0.0, -0.0, -0.0, -0.0, -0.0, -0.0, -0.0, -0.0, -0.0, -0.0, -0.0, -0.0, -0.0, -0.0, -0.0, -0.0, -0.0, -0.0, -0.0, -0.0, -0.0, -0.0, -0.0, -0.0, -0.0, -0.0, -0.0, -0.0, -0.0, -0.0, -0.0, -0.0, -0.0, -0.0, -0.0, -0.0, -0.0, -0.0, -0.0, -0.0, -0.0, -0.0, -0.0, -0.0, -0.0, -0.0, -0.0, -0.0, -0.0, -0.0, -0.0, -1.7756006070928429E-5, -1.955926027849794E-5, -2.1265642444599059E-5, -2.2878087249309936E-5, -2.4399475238503513E-5, -2.5832632877734329E-5, -2.7180332648224444E-5, -2.8445293182983732E-5, -2.9630179441154765E-5, -3.0737602918726609E-5, -3.1770121893815045E-5, -3.2730241704758869E-5, -3.3620415059333691E-5, -3.4443042373434618E-5, -3.5200472137629193E-5, -3.5895001310030509E-5, -3.652887573398812E-5, -3.7104290579141277E-5, -3.7623390804425058E-5, -3.808827164166491E-5, -3.8500979098439383E-5, -3.886351047893401E-5, -3.9177814921551905E-5, -3.9445793952087749E-5, -3.966930205131298E-5, -3.98501472358593E-5, -3.9990091651326829E-5, -4.0090852176581095E-5, -4.0154101038240283E-5, 0.0, 0.0, 0.0, 0.0, 0.0, 0.0, 0.0, 0.0, 0.0, 0.0, 0.0, 0.0, 0.0, 0.0, 0.0, 0.0, 0.0, 0.0, 0.0, 0.0, 0.0, 0.0, 0.0, 0.0, 0.0, 0.0, 0.0, 0.0, 0.0, 0.0, 0.0, 0.0, 0.0, 0.0, 0.0, 0.0, 0.0, 0.0, 0.0, 0.0, 0.0, 0.0, 0.0, 0.0, 0.0, 0.0, 0.0, 0.0, 0.0, 0.0, 0.0, 0.0, 0.0, 0.0, 0.0, 0.0, 0.0, 0.0, 0.0, 0.0, 0.0, 0.0, 0.0, 0.0, 0.0, 0.0, 0.0, 0.0, 0.0, 0.0, 0.0, 0.0, 0.0, 0.0, 0.0, 0.0, 0.0, 0.0, 0.0, 0.0, 0.0, 0.0, 0.0, 0.0, 0.0, 0.0, 0.0, 0.0, 0.0, 0.0, 0.0, 1.7756006070928429E-5, 1.955926027849794E-5, 2.1265642444599059E-5, 2.2878087249309936E-5, 2.4399475238503513E-5, 2.5832632877734329E-5, 2.7180332648224444E-5, 2.8445293182983732E-5, 2.9630179441154765E-5, 3.0737602918726609E-5, 3.1770121893815045E-5, 3.2730241704758869E-5, 3.3620415059333691E-5, 3.4443042373434618E-5, 3.5200472137629193E-5, 3.5895001310030509E-5, 3.652887573398812E-5, 3.7104290579141277E-5, 3.7623390804425058E-5, 3.808827164166491E-5, 3.8500979098439383E-5, 3.886351047893401E-5, 3.9177814921551905E-5, 3.9445793952087749E-5, 3.966930205131298E-5, 3.98501472358593E-5, 3.9990091651326829E-5, 4.0090852176581095E-5, 4.0154101038240283E-5, 0.0, 0.0, 0.0, 0.0, -0.0, -0.0, -0.0, -0.0, -0.0, -0.0, -0.0, -0.0, -0.0, -0.0, -0.0, -0.0, -0.0, -0.0, -0.0, -0.0, -0.0, -0.0, -0.0, -0.0, -0.0, -0.0, -0.0, -0.0, -0.0, -0.0, -0.0, -0.0, -0.0, -0.0, -0.0, -0.0, -0.0, -0.0, -0.0, -0.0, -0.0, -0.0, -0.0, -0.0, -0.0, -0.0, -0.0, -0.0, -0.0, -0.0, -0.0, -0.0, -0.0, -0.0, -0.0, -0.0, -0.0, -0.0, -0.0, -0.0, -0.0, -0.0, -0.0, -0.0, -0.0, -0.0, -0.0, -0.0, -0.0, -0.0, -0.0, -0.0, -0.0, -0.0, -0.0, -0.0, -0.0, -0.0, -0.0, -0.0, -0.0, -0.0, -0.0, -0.0, -0.0, -0.0, -0.0, -0.0, -0.0, -0.0, -0.0, -0.0, -0.0, -0.0, -0.0, -0.0, -0.0, -0.0, -0.0, -0.0, -0.0, -0.0, -0.0, -0.0, -0.0, -0.0, -0.0, -0.0, -0.0, -0.0, -0.0, -0.0, -0.0, -0.0, -0.0, -0.0, -0.0, -0.0, -0.0, -0.0, -0.0, -0.0, -0.0, -0.0, 0.0, 0.0, 0.0, 0.0, 0.0, 0.0, 0.0, 0.0, 0.0, 0.0, 0.0, 0.0, 0.0, 0.0, 0.0, 0.0, 0.0, 0.0, 0.0, 0.0, 0.0, 0.0, 0.0, 0.0, 0.0, 0.0, 0.0, 0.0, 0.0, 0.0, 0.0, 0.0, 0.0, 0.0, 0.0, 0.0, 0.0, 0.0, 0.0, 0.0, 0.0, 0.0, 0.0, 0.0, 0.0, 0.0, 0.0, 0.0, 0.0, 0.0, 0.0, 0.0, 0.0, 0.0, 0.0, 0.0, 0.0, 0.0, 0.0, 0.0, 0.0, 0.0, 0.0, 0.0, 0.0, 0.0, 0.0, 0.0, 0.0, 0.0, 0.0, 0.0, 0.0, 0.0, 0.0, 0.0, 0.0, 0.0, 0.0, 0.0, 0.0, 0.0, 0.0, 0.0, 0.0, 0.0, 0.0, 0.0, 0.0, 0.0, 0.0, 0.0, 0.0, 0.0, 0.0, 0.0, 0.0, 0.0, 0.0, 0.0, 0.0, 0.0, 0.0, 0.0, 0.0, 0.0, 0.0, 0.0, 0.0, 0.0, 0.0, 0.0, 0.0, 0.0, 0.0, 0.0, 0.0, 0.0, 0.0, 0.0, 0.0, 0.0, 0.0, 0.0, -0.0, -0.0, -0.0, -0.0, -0.0, -0.0, -0.0, -0.0, -0.0, -0.0, -0.0, -0.0, -0.0, -0.0, -0.0, -0.0, -0.0, -0.0, -0.0, -0.0, -0.0, -0.0, -0.0, -0.0, -0.0, -0.0, -0.0, -0.0, -0.0, -0.0, -0.0, -0.0, -0.0, -0.0, -0.0, -0.0, -0.0, -0.0, -0.0, -0.0, -0.0, -0.0, -0.0, -0.0, -0.0, -0.0, -0.0, -0.0, -0.0, -0.0, -0.0, -0.0, -0.0, -0.0, -0.0, -0.0, -0.0, -0.0, -0.0, -0.0, -0.0, -0.0, -0.0, -0.0, -0.0, -0.0, -0.0, -0.0, -0.0, -0.0, -0.0, -0.0, -0.0, -0.0, -0.0, -0.0, -0.0, -0.0, -0.0, -0.0, -0.0, -0.0, -0.0, -0.0, -0.0, -0.0, -0.0, -0.0, -0.0, -0.0, -0.0, -0.0, -1.7756006070928429E-5, -1.955926027849794E-5, -2.1265642444599059E-5, -2.2878087249309936E-5, -2.4399475238503513E-5, -2.5832632877734329E-5, -2.7180332648224444E-5, -2.8445293182983732E-5, -2.9630179441154765E-5, -3.0737602918726609E-5, -3.1770121893815045E-5, -3.2730241704758869E-5, -3.3620415059333691E-5, -3.4443042373434618E-5, -3.5200472137629193E-5, -3.5895001310030509E-5, -3.652887573398812E-5, -3.7104290579141277E-5, -3.7623390804425058E-5, -3.808827164166491E-5, -3.8500979098439383E-5, -3.886351047893401E-5, -3.9177814921551905E-5, -3.9445793952087749E-5, -3.966930205131298E-5, -3.98501472358593E-5, -3.9990091651326829E-5, -4.0090852176581095E-5, 0.0, 0.0, 0.0, 0.0, 0.0, 0.0, 0.0, 0.0, 0.0, 0.0, 0.0, 0.0, 0.0, 0.0, 0.0, 0.0, 0.0, 0.0, 0.0, 0.0, 0.0, 0.0, 0.0, 0.0, 0.0, 0.0, 0.0, 0.0, 0.0, 0.0, 0.0, 0.0, 0.0, 0.0, 0.0, 0.0, 0.0, 0.0, 0.0, 0.0, 0.0, 0.0, 0.0, 0.0, 0.0, 0.0, 0.0, 0.0, 0.0, 0.0, 0.0, 0.0, 0.0, 0.0, 0.0, 0.0, 0.0, 0.0, 0.0, 0.0, 0.0, 0.0, 0.0, 0.0, 0.0, 0.0, 0.0, 0.0, 0.0, 0.0, 0.0, 0.0, 0.0, 0.0, 0.0, 0.0, 0.0, 0.0, 0.0, 0.0, 0.0, 0.0, 0.0, 0.0, 0.0, 0.0, 0.0, 0.0, 0.0, 0.0, 0.0, 0.0, 1.7756006070928429E-5, 1.955926027849794E-5, 2.1265642444599059E-5, 2.2878087249309936E-5, 2.4399475238503513E-5, 2.5832632877734329E-5, 2.7180332648224444E-5, 2.8445293182983732E-5, 2.9630179441154765E-5, 3.0737602918726609E-5, 3.1770121893815045E-5, 3.2730241704758869E-5, 3.3620415059333691E-5, 3.4443042373434618E-5, 3.5200472137629193E-5, 3.5895001310030509E-5, 3.652887573398812E-5, 3.7104290579141277E-5, 3.7623390804425058E-5, 3.808827164166491E-5, 3.8500979098439383E-5, 3.886351047893401E-5, 3.9177814921551905E-5, 3.9445793952087749E-5, 3.966930205131298E-5, 3.98501472358593E-5, 3.9990091651326829E-5, 4.0090852176581095E-5, 0.0, 0.0, 0.0, 0.0, -0.0, -0.0, -0.0, -0.0, -0.0, -0.0, -0.0, -0.0, -0.0, -0.0, -0.0, -0.0, -0.0, -0.0, -0.0, -0.0, -0.0, -0.0, -0.0, -0.0, -0.0, -0.0, -0.0, -0.0, -0.0, -0.0, -0.0, -0.0, -0.0, -0.0, -0.0, -0.0, -0.0, -0.0, -0.0, -0.0, -0.0, -0.0, -0.0, -0.0, -0.0, -0.0, -0.0, -0.0, -0.0, -0.0, -0.0, -0.0, -0.0, -0.0, -0.0, -0.0, -0.0, -0.0, -0.0, -0.0, -0.0, -0.0, -0.0, -0.0, -0.0, -0.0, -0.0, -0.0, -0.0, -0.0, -0.0, -0.0, -0.0, -0.0, -0.0, -0.0, -0.0, -0.0, -0.0, -0.0, -0.0, -0.0, -0.0, -0.0, -0.0, -0.0, -0.0, -0.0, -0.0, -0.0, -0.0, -0.0, -0.0, -0.0, -0.0, -0.0, -0.0, -0.0, -0.0, -0.0, -0.0, -0.0, -0.0, -0.0, -0.0, -0.0, -0.0, -0.0, -0.0, -0.0, -0.0, -0.0, -0.0, -0.0, -0.0, -0.0, -0.0, -0.0, -0.0, -0.0, -0.0, -0.0, -0.0, -0.0, 0.0, 0.0, 0.0, 0.0, 0.0, 0.0, 0.0, 0.0, 0.0, 0.0, 0.0, 0.0, 0.0, 0.0, 0.0, 0.0, 0.0, 0.0, 0.0, 0.0, 0.0, 0.0, 0.0, 0.0, 0.0, 0.0, 0.0, 0.0, 0.0, 0.0, 0.0, 0.0, 0.0, 0.0, 0.0, 0.0, 0.0, 0.0, 0.0, 0.0, 0.0, 0.0, 0.0, 0.0, 0.0, 0.0, 0.0, 0.0, 0.0, 0.0, 0.0, 0.0, 0.0, 0.0, 0.0, 0.0, 0.0, 0.0, 0.0, 0.0, 0.0, 0.0, 0.0, 0.0, 0.0, 0.0, 0.0, 0.0, 0.0, 0.0, 0.0, 0.0, 0.0, 0.0, 0.0, 0.0, 0.0, 0.0, 0.0, 0.0, 0.0, 0.0, 0.0, 0.0, 0.0, 0.0, 0.0, 0.0, 0.0, 0.0, 0.0, 0.0, 0.0, 0.0, 0.0, 0.0, 0.0, 0.0, 0.0, 0.0, 0.0, 0.0, 0.0, 0.0, 0.0, 0.0, 0.0, 0.0, 0.0, 0.0, 0.0, 0.0, 0.0, 0.0, 0.0, 0.0, 0.0, 0.0, 0.0, 0.0, 0.0, 0.0, 0.0, 0.0, -0.0, -0.0, -0.0, -0.0, -0.0, -0.0, -0.0, -0.0, -0.0, -0.0, -0.0, -0.0, -0.0, -0.0, -0.0, -0.0, -0.0, -0.0, -0.0, -0.0, -0.0, -0.0, -0.0, -0.0, -0.0, -0.0, -0.0, -0.0, -0.0, -0.0, -0.0, -0.0, -0.0, -0.0, -0.0, -0.0, -0.0, -0.0, -0.0, -0.0, -0.0, -0.0, -0.0, -0.0, -0.0, -0.0, -0.0, -0.0, -0.0, -0.0, -0.0, -0.0, -0.0, -0.0, -0.0, -0.0, -0.0, -0.0, -0.0, -0.0, -0.0, -0.0, -0.0, -0.0, -0.0, -0.0, -0.0, -0.0, -0.0, -0.0, -0.0, -0.0, -0.0, -0.0, -0.0, -0.0, -0.0, -0.0, -0.0, -0.0, -0.0, -0.0, -0.0, -0.0, -0.0, -0.0, -0.0, -0.0, -0.0, -0.0, -0.0, -0.0, -0.0, -1.7756006070928429E-5, -1.955926027849794E-5, -2.1265642444599059E-5, -2.2878087249309936E-5, -2.4399475238503513E-5, -2.5832632877734329E-5, -2.7180332648224444E-5, -2.8445293182983732E-5, -2.9630179441154765E-5, -3.0737602918726609E-5, -3.1770121893815045E-5, -3.2730241704758869E-5, -3.3620415059333691E-5, -3.4443042373434618E-5, -3.5200472137629193E-5, -3.5895001310030509E-5, -3.652887573398812E-5, -3.7104290579141277E-5, -3.7623390804425058E-5, -3.808827164166491E-5, -3.8500979098439383E-5, -3.886351047893401E-5, -3.9177814921551905E-5, -3.9445793952087749E-5, -3.966930205131298E-5, -3.98501472358593E-5, -3.9990091651326829E-5, 0.0, 0.0, 0.0, 0.0, 0.0, 0.0, 0.0, 0.0, 0.0, 0.0, 0.0, 0.0, 0.0, 0.0, 0.0, 0.0, 0.0, 0.0, 0.0, 0.0, 0.0, 0.0, 0.0, 0.0, 0.0, 0.0, 0.0, 0.0, 0.0, 0.0, 0.0, 0.0, 0.0, 0.0, 0.0, 0.0, 0.0, 0.0, 0.0, 0.0, 0.0, 0.0, 0.0, 0.0, 0.0, 0.0, 0.0, 0.0, 0.0, 0.0, 0.0, 0.0, 0.0, 0.0, 0.0, 0.0, 0.0, 0.0, 0.0, 0.0, 0.0, 0.0, 0.0, 0.0, 0.0, 0.0, 0.0, 0.0, 0.0, 0.0, 0.0, 0.0, 0.0, 0.0, 0.0, 0.0, 0.0, 0.0, 0.0, 0.0, 0.0, 0.0, 0.0, 0.0, 0.0, 0.0, 0.0, 0.0, 0.0, 0.0, 0.0, 0.0, 0.0, 1.7756006070928429E-5, 1.955926027849794E-5, 2.1265642444599059E-5, 2.2878087249309936E-5, 2.4399475238503513E-5, 2.5832632877734329E-5, 2.7180332648224444E-5, 2.8445293182983732E-5, 2.9630179441154765E-5, 3.0737602918726609E-5, 3.1770121893815045E-5, 3.2730241704758869E-5, 3.3620415059333691E-5, 3.4443042373434618E-5, 3.5200472137629193E-5, 3.5895001310030509E-5, 3.652887573398812E-5, 3.7104290579141277E-5, 3.7623390804425058E-5, 3.808827164166491E-5, 3.8500979098439383E-5, 3.886351047893401E-5, 3.9177814921551905E-5, 3.9445793952087749E-5, 3.966930205131298E-5, 3.98501472358593E-5, 3.9990091651326829E-5, 0.0, 0.0, 0.0, 0.0, -0.0, -0.0, -0.0, -0.0, -0.0, -0.0, -0.0, -0.0, -0.0, -0.0, -0.0, -0.0, -0.0, -0.0, -0.0, -0.0, -0.0, -0.0, -0.0, -0.0, -0.0, -0.0, -0.0, -0.0, -0.0, -0.0, -0.0, -0.0, -0.0, -0.0, -0.0, -0.0, -0.0, -0.0, -0.0, -0.0, -0.0, -0.0, -0.0, -0.0, -0.0, -0.0, -0.0, -0.0, -0.0, -0.0, -0.0, -0.0, -0.0, -0.0, -0.0, -0.0, -0.0, -0.0, -0.0, -0.0, -0.0, -0.0, -0.0, -0.0, -0.0, -0.0, -0.0, -0.0, -0.0, -0.0, -0.0, -0.0, -0.0, -0.0, -0.0, -0.0, -0.0, -0.0, -0.0, -0.0, -0.0, -0.0, -0.0, -0.0, -0.0, -0.0, -0.0, -0.0, -0.0, -0.0, -0.0, -0.0, -0.0, -0.0, -0.0, -0.0, -0.0, -0.0, -0.0, -0.0, -0.0, -0.0, -0.0, -0.0, -0.0, -0.0, -0.0, -0.0, -0.0, -0.0, -0.0, -0.0, -0.0, -0.0, -0.0, -0.0, -0.0, -0.0, -0.0, -0.0, -0.0, -0.0, -0.0, -0.0, 0.0, 0.0, 0.0, 0.0, 0.0, 0.0, 0.0, 0.0, 0.0, 0.0, 0.0, 0.0, 0.0, 0.0, 0.0, 0.0, 0.0, 0.0, 0.0, 0.0, 0.0, 0.0, 0.0, 0.0, 0.0, 0.0, 0.0, 0.0, 0.0, 0.0, 0.0, 0.0, 0.0, 0.0, 0.0, 0.0, 0.0, 0.0, 0.0, 0.0, 0.0, 0.0, 0.0, 0.0, 0.0, 0.0, 0.0, 0.0, 0.0, 0.0, 0.0, 0.0, 0.0, 0.0, 0.0, 0.0, 0.0, 0.0, 0.0, 0.0, 0.0, 0.0, 0.0, 0.0, 0.0, 0.0, 0.0, 0.0, 0.0, 0.0, 0.0, 0.0, 0.0, 0.0, 0.0, 0.0, 0.0, 0.0, 0.0, 0.0, 0.0, 0.0, 0.0, 0.0, 0.0, 0.0, 0.0, 0.0, 0.0, 0.0, 0.0, 0.0, 0.0, 0.0, 0.0, 0.0, 0.0, 0.0, 0.0, 0.0, 0.0, 0.0, 0.0, 0.0, 0.0, 0.0, 0.0, 0.0, 0.0, 0.0, 0.0, 0.0, 0.0, 0.0, 0.0, 0.0, 0.0, 0.0, 0.0, 0.0, 0.0, 0.0, 0.0, 0.0, -0.0, -0.0, -0.0, -0.0, -0.0, -0.0, -0.0, -0.0, -0.0, -0.0, -0.0, -0.0, -0.0, -0.0, -0.0, -0.0, -0.0, -0.0, -0.0, -0.0, -0.0, -0.0, -0.0, -0.0, -0.0, -0.0, -0.0, -0.0, -0.0, -0.0, -0.0, -0.0, -0.0, -0.0, -0.0, -0.0, -0.0, -0.0, -0.0, -0.0, -0.0, -0.0, -0.0, -0.0, -0.0, -0.0, -0.0, -0.0, -0.0, -0.0, -0.0, -0.0, -0.0, -0.0, -0.0, -0.0, -0.0, -0.0, -0.0, -0.0, -0.0, -0.0, -0.0, -0.0, -0.0, -0.0, -0.0, -0.0, -0.0, -0.0, -0.0, -0.0, -0.0, -0.0, -0.0, -0.0, -0.0, -0.0, -0.0, -0.0, -0.0, -0.0, -0.0, -0.0, -0.0, -0.0, -0.0, -0.0, -0.0, -0.0, -0.0, -0.0, -0.0, -0.0, -1.7756006070928429E-5, -1.955926027849794E-5, -2.1265642444599059E-5, -2.2878087249309936E-5, -2.4399475238503513E-5, -2.5832632877734329E-5, -2.7180332648224444E-5, -2.8445293182983732E-5, -2.9630179441154765E-5, -3.0737602918726609E-5, -3.1770121893815045E-5, -3.2730241704758869E-5, -3.3620415059333691E-5, -3.4443042373434618E-5, -3.5200472137629193E-5, -3.5895001310030509E-5, -3.652887573398812E-5, -3.7104290579141277E-5, -3.7623390804425058E-5, -3.808827164166491E-5, -3.8500979098439383E-5, -3.886351047893401E-5, -3.9177814921551905E-5, -3.9445793952087749E-5, -3.966930205131298E-5, -3.98501472358593E-5, 0.0, 0.0, 0.0, 0.0, 0.0, 0.0, 0.0, 0.0, 0.0, 0.0, 0.0, 0.0, 0.0, 0.0, 0.0, 0.0, 0.0, 0.0, 0.0, 0.0, 0.0, 0.0, 0.0, 0.0, 0.0, 0.0, 0.0, 0.0, 0.0, 0.0, 0.0, 0.0, 0.0, 0.0, 0.0, 0.0, 0.0, 0.0, 0.0, 0.0, 0.0, 0.0, 0.0, 0.0, 0.0, 0.0, 0.0, 0.0, 0.0, 0.0, 0.0, 0.0, 0.0, 0.0, 0.0, 0.0, 0.0, 0.0, 0.0, 0.0, 0.0, 0.0, 0.0, 0.0, 0.0, 0.0, 0.0, 0.0, 0.0, 0.0, 0.0, 0.0, 0.0, 0.0, 0.0, 0.0, 0.0, 0.0, 0.0, 0.0, 0.0, 0.0, 0.0, 0.0, 0.0, 0.0, 0.0, 0.0, 0.0, 0.0, 0.0, 0.0, 0.0, 0.0, 1.7756006070928429E-5, 1.955926027849794E-5, 2.1265642444599059E-5, 2.2878087249309936E-5, 2.4399475238503513E-5, 2.5832632877734329E-5, 2.7180332648224444E-5, 2.8445293182983732E-5, 2.9630179441154765E-5, 3.0737602918726609E-5, 3.1770121893815045E-5, 3.2730241704758869E-5, 3.3620415059333691E-5, 3.4443042373434618E-5, 3.5200472137629193E-5, 3.5895001310030509E-5, 3.652887573398812E-5, 3.7104290579141277E-5, 3.7623390804425058E-5, 3.808827164166491E-5, 3.8500979098439383E-5, 3.886351047893401E-5, 3.9177814921551905E-5, 3.9445793952087749E-5, 3.966930205131298E-5, 3.98501472358593E-5, 0.0, 0.0, 0.0, 0.0, -0.0, -0.0, -0.0, -0.0, -0.0, -0.0, -0.0, -0.0, -0.0, -0.0, -0.0, -0.0, -0.0, -0.0, -0.0, -0.0, -0.0, -0.0, -0.0, -0.0, -0.0, -0.0, -0.0, -0.0, -0.0, -0.0, -0.0, -0.0, -0.0, -0.0, -0.0, -0.0, -0.0, -0.0, -0.0, -0.0, -0.0, -0.0, -0.0, -0.0, -0.0, -0.0